(* IEC 61131-3 sources: plcassist-cli/packages/volt-lsp-iec/test-corpus/pro2193/Device/Plc Logic/Application/09 Misc/Library Manager/L_TS2P_TechModulesSynchronizingCamming (part 2) *)

(* ---- L_TS2P_SYNCANDCORRECTIONSTATE.fb ---- *)
FUNCTION_BLOCK L_TS2P_SYNCANDCORRECTIONSTATE EXTENDS L_TB2P_TechModuleBase
VAR_INPUT
	XUSEORIGINAL : BOOL;
	XENABLE : BOOL;
	XENABLEOPERATION : BOOL;
	XRESETERROR : BOOL;
	XQSPAPPLICATION : BOOL;
	XABORT : BOOL;
	XJOGPOS : BOOL;
	XJOGNEG : BOOL;
	XHOMEEXECUTE : BOOL;
	LROVERRIDE : LREAL := 1;
	SCCTRLBASICMOTION : L_TB2P_scCtrlBasicMotion;
	SCPAR : L_TS2P_scPar_SyncAndCorrectionState;
	SCACCESSPOINTS : L_TS2P_scAP_SyncAndCorrectionState;
	MASTERVALUES : L_MC1P_IAXIS_REF_MASTERVALUES;
	XSYNCIN : BOOL;
	XSYNCPOSRESTORE : BOOL;
	LRSETBASEVEL : LREAL;
	LRSETOFFSETPOS : LREAL;
	XTRIMPOS : BOOL;
	XTRIMNEG : BOOL;
	XTRIMRESET : BOOL;
	SCTPRECDATA_MARKSENSOR : L_MC1P_TpReceiveData;
	SCTPRECDATA_TOOLSENSOR : L_MC1P_TpReceiveData;
	XTEACHMARKWINDOW : BOOL;
	XTEACHMARKWINDOWTOOL : BOOL;
	XGEARFACTORCORR : BOOL;
	XGEARFACTORCORRHOLD : BOOL;
END_VAR
VAR_OUTPUT
	XREADYFOROPERATION : BOOL;
	XOPERATIONENABLED : BOOL;
	XREADYFORMOTION : BOOL;
	XERROR : BOOL;
	XWARNING : BOOL;
	EERRORID : L_IE1P_Error;
	XSTOACTIVE : BOOL;
	XQSPACTIVE : BOOL;
	XABORTBUSY : BOOL;
	XABORTDONE : BOOL;
	XJOGGINGBUSY : BOOL;
	XHOMINGBUSY : BOOL;
	XHOMINGDONE : BOOL;
	XISHOMED : BOOL;
	ETMSTATE : L_TB2P_States := L_TB2P_States.DISABLED;
	SCSTATUSBASICMOTION : L_TB2P_scStatusBasicMotion;
	LRACTVEL : LREAL;
	LRSETVELOUT : LREAL;
	LRACTPOS : LREAL;
	LRSETPOSOUT : LREAL;
	LRACTFOLLOWINGERROR : LREAL;
	SCSIGNALFLOW : L_TS2P_scSF_SyncAndCorrectionState;
	XSYNCHRONISED : BOOL;
	XACCDECSYNC : BOOL;
	XOFFSETTRIMACTIVE : BOOL;
	XBASEVELOCITYACTIVE : BOOL;
	LROFFSETTOTAL : LREAL;
	LRSETMARKCORROUT : LREAL;
	XMARKWINDOWTEACHED : BOOL;
	LRGEARFACTORCORR : LREAL;
	LRSETTOOLCORROUT : LREAL;
	XMARKWINDOWTEACHEDTOOL : BOOL;
END_VAR
VAR_IN_OUT
	AXIS : AXIS_REF;
END_VAR
VAR
	XINTERNALCONTROL : BOOL;
	XINTERNALCONTROLACTIVE : BOOL;
	XINTERNALCONTROLACTIVE_OLD : BOOL;
	ITFCONNECTORSYNCANDCORRECTION : L_TS2P_IConnectorSyncAndCorrection;
	TM_INT : L_TS2P_TM_SyncAndCorrectionState;
	SCPAR_INT : L_TS2P_scPar_SyncAndCorrectionState;
	XSYNCIN_INT : BOOL;
	XSYNCPOSRESTORE_INT : BOOL;
	LRSETBASEVEL_INT : LREAL;
	LRSETOFFSETPOS_INT : LREAL;
	XTRIMPOS_INT : BOOL;
	XTRIMNEG_INT : BOOL;
	XTRIMRESET_INT : BOOL;
	XTEACHMARKWINDOW_INT : BOOL;
	XTEACHMARKWINDOWTOOL_INT : BOOL;
	XGEARFACTORCORR_INT : BOOL;
	XGEARFACTORCORRHOLD_INT : BOOL;
	XUSEORIGINAL_OLD : BOOL;
	ITFBASICMOTIONBASE : L_TB2P.L_TB2P_IBasicMotionBase;
	ITFITECHMODULEINTERNAL : L_TB2P_ITechModuleInternal;
	ITFSYNCANDCORRECTIONEXTENSION : L_TS2P_ISyncAndCorrectionState;
	ITFSYNCPOSEXTENSION : L_TS2P_ISyncPosBase;
	LRJERKDEC : LREAL;
	LRJOGGINGJERKDEC : LREAL;
	REMAININGTIMEOFPROFILE : LREAL;
	REMAININGTIMEOFPROFILEAVAILABLE : BOOL;
END_VAR
END_FUNCTION_BLOCK

METHOD GET_PAP : POINTER TO L_TB2P_scAP_TM_MotionControl
END_METHOD

METHOD GET_PPAR : POINTER TO L_TB2P.L_TB2P_scPar_TM_MotionControl
END_METHOD

METHOD GET_PSF : POINTER TO L_TB2P_scSF_TM_MotionControl
END_METHOD

METHOD CALL_ABC
VAR_INPUT
	ITFTECHMODULE : L_TB2P.L_TB2P_IBasicMotionBase;
	XQSPAPPLICATION : BOOL;
	XHALT : BOOL;
	XABORT : BOOL;
	XHOMEEXECUTE : BOOL;
	XJOGPOS : BOOL;
	XJOGNEG : BOOL;
	XFINISHPOSITIONING : BOOL;
	XMOVEVELEXECUTE : BOOL;
	XMOVEABSEXECUTE : BOOL;
	XMOVERELEXECUTE : BOOL;
	XENABLEOPERATION : BOOL;
	XRESETERROR : BOOL;
	XENABLEPOSITIVE : BOOL;
	XENABLENEGATIVE : BOOL;
	XDISABLESWLIMIT : BOOL;
	LROVERRIDE : LREAL;
	LROVERRIDEACC : LREAL;
	LROVERRIDEJERK : LREAL;
	XRESETHOMEPOSITION : BOOL;
	XCONTINUOUSUPDATE : BOOL;
	LRPOS_DIST : LREAL;
	LRVEL : LREAL;
	LRACC : LREAL;
	LRDEC : LREAL;
	LRJERK : LREAL;
	EDIRECTION : L_TB2P.MC_DIRECTION;
	SCHOMEEXTTP : L_TB2P.MC_TRIGGER_REF;
	XHOMEABSSWITCH : BOOL;
	XSPECIALABORTBEHAVIOR : BOOL;
	LRABORTDEC : LREAL;
	LRABORTJERK : LREAL;
END_VAR
VAR_OUTPUT
	XERROR : BOOL;
	EERRORID : L_TB2P.L_IE1P_Error;
	XFUNBUSY : BOOL;
	XFUNDONE : BOOL;
	XFUNCOMMANDABORTED : BOOL;
	EFUNSTATEACT : L_TB2P.L_MC1P_ABC_State;
	ECONTROLMODE : L_TB2P.L_MC1P_ControlMode;
	XISHOMED : BOOL;
	XHWLIMITSWITCHNEG : BOOL;
	XHWLIMITSWITCHPOS : BOOL;
	XSWLIMITENABLED : BOOL;
	XSWLIMITSWITCHNEG : BOOL;
	XSWLIMITSWITCHPOS : BOOL;
	EAXISTYPE : L_TB2P.L_MC1P_DriveType;
	EAXISSTATE : L_TB2P.L_MC1P_AXIS_STATE;
	XSTOACTIVE : BOOL;
	XREADYFOROPERATION : BOOL;
	XOPERATIONENABLED : BOOL;
	XREADYFORMOTION : BOOL;
	XAXISWARNING : BOOL;
	XAXISERROR : BOOL;
	EAXISERRORID : L_TB2P.L_IE1P_Error;
	XDRIVEWARNING : BOOL;
	XDRIVEERROR : BOOL;
	DWDRIVEERRORID : DWORD;
	LRACTPOS : LREAL;
	LRACTVEL : LREAL;
	LRSETPOSOUT : LREAL;
	LRSETVELOUT : LREAL;
	LRACTFOLLOWINGERROR : LREAL;
	XINPOSITION : BOOL;
	XSTANDSTILLSETVELOCITY : BOOL;
	XSTANDSTILLACTVELOCITY : BOOL;
	XCONSTANTVELOCITY : BOOL;
	XACCELERATING : BOOL;
	XDECELERATING : BOOL;
	XDIRECTIONPOSITIVE : BOOL;
	XDIRECTIONNEGATIVE : BOOL;
	XAXISAVAILABLE : BOOL;
END_VAR
VAR_IN_OUT
	AXIS : AXIS_REF;
END_VAR
END_METHOD

METHOD ADDOFFSET
VAR_INPUT
	ITFTECHMODULE : L_TS2P_ISyncPosBase;
	LRSETPOS : LREAL;
	LRSETVEL : LREAL;
	LRSETOFFSET : LREAL;
	LRSETOFFSETVEL : LREAL;
	ETRAVERSINGRANGE : L_MC1P.L_MC1P_TraversingRange;
	LRCYCLELENGTH : LREAL;
END_VAR
VAR_OUTPUT
	XERROR : BOOL;
	EERRORID : L_IE1P.L_IE1P_Error;
	LRSETPOSOUT : LREAL;
	LRSETVELOUT : LREAL;
END_VAR
END_METHOD

METHOD CLUTCH
VAR_INPUT
	ITFTECHMODULE : L_TS2P_ISyncPosBase;
	XENABLE : BOOL;
	XSYNCIN : BOOL;
	LRSETBASEVELOCITY : LREAL;
	ESYNCMODE : L_TB2P_SyncMode;
	EALLOWEDDIRECTION : L_TB2P_AllowedDirection;
	LRSYNCVEL : LREAL;
	LRSYNCACC : LREAL;
	LRSYNCDEC : LREAL;
	LRSYNCJERK : LREAL;
	LRSYNCINDIST : LREAL;
	LRSYNCOUTDIST : LREAL;
	LRSYNCOUTPOS : LREAL;
	XLOADCLUTCHOFFSET : BOOL;
	LRLOADCLUTCHOFFSET : LREAL;
	LRCYCLICMASTERPOS : LREAL;
	LRCYCLICMASTERVEL : LREAL;
	ETRAVERSINGRANGEMASTER : L_MC1P_TraversingRange;
	LRCYCLELENGTHMASTER : LREAL;
	LRCYCLICAXISPOS : LREAL;
	LRCYCLICAXISVEL : LREAL;
	LRCYCLICAXISACC : LREAL;
	ETRAVERSINGRANGEAXIS : L_MC1P_TraversingRange;
	LRCYCLELENGTHAXIS : LREAL;
END_VAR
VAR_OUTPUT
	XERROR : BOOL;
	EERRORID : L_IE1P.L_IE1P_Error;
	XBUSY : BOOL;
	XDONE : BOOL;
	XSYNCHRONISED : BOOL;
	XACCDECSYNC : BOOL;
	XINBASEVELOCITY : BOOL;
	LRSETPOSOUT : LREAL;
	LRSETVELOUT : LREAL;
	LRSETACCOUT : LREAL;
	LRCLUTCHOFFSETOUT : LREAL;
END_VAR
END_METHOD

METHOD GEARBOX
VAR_INPUT
	ITFTECHMODULE : L_TS2P_ISyncPosBase;
	XENABLE : BOOL;
	LRSETPOSX : LREAL;
	LRSETVELX : LREAL;
	DWNUMERATOR : DWORD;
	DWDENOMINATOR : DWORD;
	LRCYCLELENGTHX : LREAL;
	LRCYCLELENGTHY : LREAL;
	ETRAVERSINGRANGEX : L_MC1P.L_MC1P_TraversingRange;
	ETRAVERSINGRANGEY : L_MC1P.L_MC1P_TraversingRange;
	XLOADGEARBOXPOS : BOOL;
	LRLOADGEARBOXPOS : LREAL;
END_VAR
VAR_OUTPUT
	XERROR : BOOL;
	EERRORID : L_IE1P.L_IE1P_Error;
	LRSETPOSOUT : LREAL;
	LRSETVELOUT : LREAL;
END_VAR
END_METHOD

METHOD OFFSETANDTRIM
VAR_INPUT
	ITFTECHMODULE : L_TS2P_ISyncPosBase;
	XENABLE : BOOL;
	LRSETOFFSET : LREAL;
	XTRIMPOS : BOOL;
	XTRIMNEG : BOOL;
	LRSETTRIMDISTANCE : LREAL;
	ETRIMMODE : L_TS2P_TrimMode;
	XLOADOFFSET : BOOL;
	XRESETTRIMOFFSET : BOOL;
	LRSETVEL : LREAL;
	LRSETACC : LREAL;
	LRSETDEC : LREAL;
	LRSETJERK : LREAL;
	WACTDIRECTION : WORD;
	EALLOWEDDIRECTION : L_TB2P.L_TB2P_AllowedDirection;
	LRCYCMASTERPOS : LREAL;
	LRCYCMASTERVEL : LREAL;
	LRCYCMASTERACC : LREAL;
END_VAR
VAR_OUTPUT
	XERROR : BOOL;
	EERRORID : L_IE1P.L_IE1P_Error;
	XBUSY : BOOL;
	XDONE : BOOL;
	LRSETOFFSETOUTTOTAL : LREAL;
	LRSETOFFSETOUTTOTALVEL : LREAL;
	LRSETOFFSETOUT : LREAL;
	LRSETOFFSETOUTTRIM : LREAL;
END_VAR
END_METHOD

METHOD FB_INIT : BOOL
VAR_INPUT
	BINITRETAINS : BOOL;
	BINCOPYCODE : BOOL;
END_VAR
END_METHOD

METHOD CALL_INTERNALCTRL
END_METHOD

(* ---- L_TS2P_SYNCANDCORRECTIONSTATE_V2.fb ---- *)
FUNCTION_BLOCK L_TS2P_SYNCANDCORRECTIONSTATE_V2 EXTENDS L_TB2P_TechModuleBase
VAR_INPUT
	XENABLE : BOOL;
	XENABLEOPERATION : BOOL;
	XRESETERROR : BOOL;
	XQSPAPPLICATION : BOOL;
	XABORT : BOOL;
	XJOGPOS : BOOL;
	XJOGNEG : BOOL;
	XHOMEEXECUTE : BOOL;
	LROVERRIDE : LREAL := 1;
	SCCTRLBASICMOTION : L_TB2P_scCtrlBasicMotion;
	SCPAR : L_TS2P_scPar_SyncAndCorrectionState;
	SCACCESSPOINTS : L_TS2P_scAP_SyncAndCorrectionState;
	MASTERVALUES : L_MC1P_IAXIS_REF_MASTERVALUES;
	XSYNCIN : BOOL;
	XSYNCPOSRESTORE : BOOL;
	LRSETBASEVEL : LREAL;
	LRSETOFFSETPOS : LREAL;
	XTRIMPOS : BOOL;
	XTRIMNEG : BOOL;
	XTRIMRESET : BOOL;
	SCTPRECDATA_MARKSENSOR : L_MC1P_TpReceiveData;
	SCTPRECDATA_TOOLSENSOR : L_MC1P_TpReceiveData;
	XTEACHMARKWINDOW : BOOL;
	XTEACHMARKWINDOWTOOL : BOOL;
	XGEARFACTORCORR : BOOL;
	XGEARFACTORCORRHOLD : BOOL;
END_VAR
VAR_OUTPUT
	XREADYFOROPERATION : BOOL;
	XOPERATIONENABLED : BOOL;
	XREADYFORMOTION : BOOL;
	XERROR : BOOL;
	XWARNING : BOOL;
	EERRORID : L_IE1P_Error;
	XSTOACTIVE : BOOL;
	XQSPACTIVE : BOOL;
	XABORTBUSY : BOOL;
	XABORTDONE : BOOL;
	XJOGGINGBUSY : BOOL;
	XHOMINGBUSY : BOOL;
	XHOMINGDONE : BOOL;
	XISHOMED : BOOL;
	ETMSTATE : L_TB2P_States := L_TB2P_States.DISABLED;
	SCSTATUSBASICMOTION : L_TB2P_scStatusBasicMotion;
	LRACTVEL : LREAL;
	LRSETVELOUT : LREAL;
	LRACTPOS : LREAL;
	LRSETPOSOUT : LREAL;
	LRACTFOLLOWINGERROR : LREAL;
	SCSIGNALFLOW : L_TS2P_scSF_SyncAndCorrectionState;
	XSYNCHRONISED : BOOL;
	XACCDECSYNC : BOOL;
	XOFFSETTRIMACTIVE : BOOL;
	XBASEVELOCITYACTIVE : BOOL;
	LROFFSETTOTAL : LREAL;
	LRSETMARKCORROUT : LREAL;
	XMARKWINDOWTEACHED : BOOL;
	LRGEARFACTORCORR : LREAL;
	LRSETTOOLCORROUT : LREAL;
	XMARKWINDOWTEACHEDTOOL : BOOL;
END_VAR
VAR_IN_OUT
	AXIS : AXIS_REF;
END_VAR
VAR
	TM_INT : L_TS2P_TM_SyncAndCorrectionState_V2 := STRUCT(ModuleHandler := ModuleHandler);
	PPAR : POINTER TO L_TS2P_scPar_SyncAndCorrectionState;
	PPAR_INT : POINTER TO L_TS2P_scPar_SyncAndCorrectionState;
	LRJERKDEC : LREAL;
	LRJOGGINGJERKDEC : LREAL;
END_VAR
END_FUNCTION_BLOCK

(* ---- L_TS2P_SYNCDRIVEPOS.fb ---- *)
FUNCTION_BLOCK L_TS2P_SYNCDRIVEPOS
VAR_INPUT
	MASTERAXIS : POINTER TO L_MC1P_IAXIS_REF_MASTERVALUES;
	XENABLE : BOOL;
	DWNUMERATOR : DWORD := 1;
	DWDENOMINATOR : DWORD := 1;
	XSYNCIN : BOOL;
	XSYNCOUTINSTANT : BOOL;
	XSYNCINSTANT : BOOL;
	XCLUTCHRELATIVE : BOOL;
	XSYNCPOSRESTORE : BOOL;
	LRSLAVESYNCOUTPOS : LREAL;
	LRSLAVESYNCINDIST : LREAL := 90;
	LRSLAVESYNCOUTDIST : LREAL := 90;
	LRSYNCOUTINSTANTDEC : LREAL := 10000;
	EALLOWEDDIRECTION : L_TB2P_AllowedDirection := L_TB2P_AllowedDirection.both;
	ESYNCMODE : L_TB2P_SyncMode := L_TB2P_SyncMode.ProfGenAbsolute;
	LRSYNCVEL : LREAL := 100;
	LRSYNCACC : LREAL := 1000.0;
	LRSYNCDEC : LREAL := 1000.0;
	LRSYNCJERK : LREAL := 10000000000.0;
	LRSETBASEVELOCITY : LREAL := 0;
	XLOADCLUTCHOFFSET : BOOL := FALSE;
	LRLOADCLUTCHOFFSET : LREAL := 0;
	XTRIMVELOCITYX : BOOL;
	XTRIMVELOCITYY : BOOL;
	LRSETTRIMDISTANCEX : LREAL := 1;
	LRSETTRIMDISTANCEY : LREAL := 1;
	XTRIMPOSX : BOOL;
	XTRIMNEGX : BOOL;
	XTRIMPOSY : BOOL;
	XTRIMNEGY : BOOL;
	XRESETTRIMX : BOOL;
	XRESETTRIMY : BOOL;
	LRSETOFFSETX : LREAL := 0;
	LRSETOFFSETTRIMVELX : LREAL := 10.0;
	LRSETOFFSETTRIMACCX : LREAL := 100.0;
	LRSETOFFSETTRIMDECX : LREAL := 100.0;
	LRSETOFFSETTRIMJERKX : LREAL := 10000.0;
	XLOADOFFSETX : BOOL;
	LRSETOFFSETY : LREAL := 0;
	LRSETOFFSETTRIMVELY : LREAL := 10.0;
	LRSETOFFSETTRIMACCY : LREAL := 100.0;
	LRSETOFFSETTRIMDECY : LREAL := 100.0;
	LRSETOFFSETTRIMJERKY : LREAL := 10000.0;
	XLOADOFFSETY : BOOL;
	XLOADSTARTSLAVEPOS : BOOL := FALSE;
	LRSTARTSLAVEPOS : LREAL;
	XLOADGEARBOXPOS : BOOL;
	LRLOADGEARBOXPOS : LREAL;
	XOPERATIONENABLED : BOOL;
END_VAR
VAR_OUTPUT
	XERROR : BOOL;
	XWARNING : BOOL;
	EERRORID : L_IE1P_Error;
	XBUSY : BOOL;
	LRSETSLAVEPOSOUT : LREAL;
	LRSETSLAVEVELOUT : LREAL;
	LRSETSLAVEACCOUT : LREAL;
	LRSETGEARBOXPOSOUT : LREAL;
	XSYNCOUTDONE : BOOL;
	XSYNCHRONISED : BOOL;
	XACCDECSYNC : BOOL;
	XOFFSETTRIMBUSY : BOOL;
	LROFFSETOUTTOTALVELX : LREAL;
	LROFFSETOUTTOTALVELY : LREAL;
	LROFFSETOUTTRIMX : LREAL;
	LROFFSETOUTTRIMY : LREAL;
	LROFFSETOUTX : LREAL;
	LROFFSETOUTY : LREAL;
	LROFFSETOUTTOTALX : LREAL;
	LROFFSETOUTTOTALY : LREAL;
	LRSETCLUTCHPOS : LREAL;
	LRSETCLUTCHVEL : LREAL;
	LRSETCLUTCHACC : LREAL;
	XBASEVELSYNCHRONISED : BOOL;
	XACCDECBASEVEL : BOOL;
	LROFFSETSYNCPOS : LREAL;
END_VAR
VAR_IN_OUT
	SLAVEAXIS : AXIS_REF;
END_VAR
VAR
	FB_GEARBOXPOSITION : L_MB1P_GearboxPositionInput;
	FB_CLUTCHEXTENDEDBASE : L_TB2P_ClutchExtendedBase;
	FB_AXISCONVERTER : L_MC2P.L_MC2P_AxisConverterBase;
	FB_OFFSETANDTRIMX : L_TS2P_OffsetAndTrim;
	FB_ADDOFFSETCYCLICX : L_MC1P_AddOffsetCyclic;
	FB_OFFSETANDTRIMY : L_TS2P_OffsetAndTrim;
	FB_ADDOFFSETCYCLICY : L_MC1P_AddOffsetCyclic;
	FB_SYNCPOSRESTOREOFFSET : L_TS2P_OffsetAndTrim;
	FB_DIRECTION : L_MC1P_GetDirection;
	LRSETOFFSETMASTER_INT : LREAL;
	LRTRIMDIST_INT : LREAL;
	XTRIMPOS_OLD : BOOL;
	XTRIMNEG_OLD : BOOL;
	XTRIMVEL : BOOL;
	LRTRIMOFFSETDIST : LREAL;
	LRLOADOFFSETMASTER_INT : LREAL := 0;
	LRLOADGEARBOXPOS_INT : LREAL;
	LRSETGEARBOXPOSOUT_INT : LREAL;
	XSETDISABLECLUTCH_INT : BOOL;
	LRLOADTRIMOFFSET_INT : LREAL := 0;
	LRSYNCOUTINSTANTDEC_INT : LREAL := 100000;
	LRSETINTEGRATETRIMVELPOSOUT_INT : LREAL;
	XSYNCPOS_OLD : BOOL;
	XRESETTRIM_OLD : BOOL;
	LRLOADOFFSET_INT : LREAL := 0;
	XSYNCINSTANT_OLD : BOOL;
	XENABLEGEARBOX : BOOL;
	LRSYNCOFFSET : LREAL;
	LRSCALING_INT : LREAL := 1;
	LRGEARBOXSTARTPOSOUT_INT : LREAL;
	DWDENOMINATOR_INT : DWORD := 1;
	XENABLE_OLD : BOOL;
	WAXESMODE : WORD;
	WAXESMODEOLD : WORD;
	LRADDOFFSETPOSOUTY_OLD : LREAL;
	LRADDOFFSETVELOUTY : LREAL;
	LRSETGEARBOXPOSOUTOLD_INT : LREAL;
	LRSETGEARBOXPOSOUTVEL_INT : LREAL;
	LRGETGEARBOXVELIN : LREAL;
	LRGETGEARBOXPOSOUT : LREAL;
	LRGETGEARBOXPOSIN : LREAL;
	LRTASKCYCLE : LREAL;
	XINIT : BOOL := TRUE;
	XCLUTCHDONE_OLD : BOOL;
	XENABLEOLD : BOOL;
	LRSETOFFSETOUTTOTALVELOLD : LREAL;
	SET_AP_LRMASTERVELSTANDSTILLDEADBAND : LREAL;
END_VAR
END_FUNCTION_BLOCK

METHOD CALL_AXESMODE
END_METHOD

METHOD CALL_CALCGEARBOXOUTVELACC
VAR_IN_OUT
	SLAVEAXIS : AXIS_REF;
END_VAR
END_METHOD

METHOD CALL_ERRORHANDLER
END_METHOD

METHOD CALL_FBMETHODS
END_METHOD

METHOD CALL_FBMETHODS_FMDISABLE
END_METHOD

METHOD CALL_FB_ADDOFFSETCYCLICX
END_METHOD

METHOD CALL_FB_ADDOFFSETCYCLICX_INPUT
END_METHOD

METHOD CALL_FB_ADDOFFSETCYCLICY
END_METHOD

METHOD CALL_FB_ADDOFFSETCYCLICY_INPUT
END_METHOD

METHOD CALL_FB_AXISCONVERTER
END_METHOD

METHOD CALL_FB_AXISCONVERTER_INPUT
END_METHOD

METHOD CALL_FB_CLUTCHEXTENDEDBASE
END_METHOD

METHOD CALL_FB_CLUTCHEXTENDEDBASE_INPUT
END_METHOD

METHOD CALL_FB_CLUTCHEXTENDEDBASE_INPUTMASTER
END_METHOD

METHOD CALL_FB_CLUTCHEXTENDEDBASE_INPUTSLAVE
VAR_IN_OUT
	SLAVEAXIS : AXIS_REF;
END_VAR
END_METHOD

METHOD CALL_FB_GEARBOXPOSITION
END_METHOD

METHOD CALL_FB_GEARBOXPOSITION_INPUT
END_METHOD

METHOD CALL_FB_GEARBOXPOSITION_LOADGEARBOXPOS
END_METHOD

METHOD CALL_FB_SYNCPOSRESTOREOFFSET
END_METHOD

METHOD CALL_FB_SYNCPOSRESTOREOFFSET_INPUT
VAR_IN_OUT
	SLAVEAXIS : AXIS_REF;
END_VAR
END_METHOD

METHOD CALL_LOADSLAVESTARTPOS
END_METHOD

METHOD CALL_OFFSETANDTRIMX
END_METHOD

METHOD CALL_OFFSETANDTRIMX_INPUT
END_METHOD

METHOD CALL_OFFSETANDTRIMY
END_METHOD

METHOD CALL_OFFSETANDTRIMY_INPUT
END_METHOD

METHOD CALL_OUTPUT
END_METHOD

METHOD CALL_OUTPUT_CLUTCHSTATE
END_METHOD

METHOD CALL_OUTPUT_OFFSET
END_METHOD

METHOD CALL_RESETCOMMANDS
END_METHOD

METHOD CALL_INIT
VAR_IN_OUT
	SLAVEAXIS : AXIS_REF;
END_VAR
END_METHOD

METHOD GET_DIRECTION
END_METHOD

METHOD GET_GETGEARBOXPOSIN : LREAL
END_METHOD

METHOD GET_GETGEARBOXPOSOUT : LREAL
END_METHOD

METHOD GET_GETGEARBOXVELIN : LREAL
END_METHOD

METHOD GET_GETGEARBOXVELOUT : LREAL
END_METHOD

METHOD GET_LRCLUTCHPOSIN : LREAL
END_METHOD

METHOD GET_LROFFSETADDOFFSETCYCLIC : LREAL
END_METHOD

METHOD SETDISABLECLUTCH : BOOL
VAR_INPUT
	XSETDISABLECLUTCH : BOOL;
END_VAR
END_METHOD

(* ---- L_TS2P_SYNCDRIVEVEL.fb ---- *)
FUNCTION_BLOCK L_TS2P_SYNCDRIVEVEL
VAR_INPUT
	MASTERAXIS : POINTER TO L_MC1P_IAXIS_REF_MASTERVALUES;
	XENABLE : BOOL;
	LRCOUPLINGX : LREAL := 1.0;
	LRCOUPLINGY : LREAL := 1.0;
	XINVERTGEARFACTOR : BOOL;
	XDISABLETOLERANCEINVERTGEARFACTOR : BOOL;
	LRTOLERANCEINVERTGEARFACTOR : LREAL := 0;
	XSYNCIN : BOOL;
	XSYNCOUTINSTANT : BOOL;
	LRSYNCACC : LREAL := 10.0;
	LRSYNCDEC : LREAL := 10.0;
	LRSYNCOUTINSTANTDEC : LREAL := 100.0;
	LRSYNCJERK : LREAL := 1.0;
	XAVOIDVELGAPS : BOOL;
	LRSETOFFSETVEL : LREAL;
	DWMODE : DWORD := 1;
	XTRIMVELOCITYX : BOOL;
	XTRIMVELOCITYY : BOOL;
	LRSETTRIMDISTANCEX : LREAL := 1;
	LRSETTRIMDISTANCEY : LREAL := 1;
	XTRIMPOSX : BOOL;
	XTRIMNEGX : BOOL;
	XTRIMPOSY : BOOL;
	XTRIMNEGY : BOOL;
	XRESETTRIMX : BOOL;
	XRESETTRIMY : BOOL;
	XSYNCVELRESET : BOOL;
	LRSETOFFSETX : LREAL := 0;
	LRSETOFFSETTRIMVELX : LREAL := 10.0;
	LRSETOFFSETTRIMACCX : LREAL := 100.0;
	LRSETOFFSETTRIMDECX : LREAL := 100.0;
	LRSETOFFSETTRIMJERKX : LREAL := 10000.0;
	XLOADOFFSETX : BOOL;
	LRSETOFFSETY : LREAL := 0;
	LRSETOFFSETTRIMVELY : LREAL := 10.0;
	LRSETOFFSETTRIMACCY : LREAL := 100.0;
	LRSETOFFSETTRIMDECY : LREAL := 100.0;
	LRSETOFFSETTRIMJERKY : LREAL := 10000.0;
	XLOADOFFSETY : BOOL;
	EALLOWEDDIRECTION : L_TB2P_AllowedDirection;
	XLOADOFFSET : BOOL;
	XLOADGROUNDVEL : BOOL;
	LRSETGROUNDVEL : LREAL;
	LRGROUNDVELACC : LREAL := 10.0;
	LRGROUNDVELDEC : LREAL := 10.0;
	LRGROUNDVELJERK : LREAL := 1.0;
END_VAR
VAR_OUTPUT
	XERROR : BOOL;
	XWARNING : BOOL;
	EERRORID : L_IE1P_Error;
	XBUSY : BOOL;
	LRSETSLAVEVELOUT : LREAL;
	LRSETSLAVEACCOUT : LREAL;
	XSYNCOUTDONE : BOOL;
	XSYNCHRONISED : BOOL;
	XACCDECSYNC : BOOL;
	XOFFSETTRIMBUSY : BOOL;
	LRPOSOFFSETOUTTRIMX : LREAL;
	LRPOSOFFSETOUTTRIMY : LREAL;
	LRPOSOFFSETOUTX : LREAL;
	LRPOSOFFSETOUTY : LREAL;
	LRPOSOFFSETOUTVELX : LREAL;
	LRVELOFFSET : LREAL;
	LROFFSETOUTTOTALX : LREAL;
	LROFFSETOUTTOTALY : LREAL;
	LROFFSETOUTTOTALVELX : LREAL;
	LROFFSETOUTTOTALVELY : LREAL;
	XBASEVELSYNCHRONISED : BOOL;
	XACCDECBASEVEL : BOOL;
	XBASEVELSYNCOUTDONE : BOOL;
	XINVERTGEARFACTORACTIVE : BOOL;
END_VAR
VAR_IN_OUT
	SLAVEAXIS : AXIS_REF;
END_VAR
VAR
	XENABLE_OLD : BOOL;
	ESTATE : L_TF1P_States := L_TF1P_States.INIT;
	ESTATE_OLD : L_TF1P_States := L_TF1P_States.INIT;
	XSTATEENTRY : BOOL;
	FB_CONVAXISV : L_MC2P_ConvAxisV;
	FB_INVERTGEARFACTOR : L_TS2P_InvertGearfactor;
	XACCDECSYNC_OLD : BOOL;
	XSYNCVEL_OLD : BOOL;
	XOPEN_OLD : BOOL;
	LRSETVELTRIM : LREAL;
	XSETDISABLECLUTCH_INT : BOOL;
	SETPOSITIONFORSYNCOLD : LREAL := 0;
	XINITFB_CLUTCHV : BOOL;
	FB_CLUTCHV : L_MC2P_ClutchVelocity;
	XINVERTGEARFACTORACTIVE_OLD : BOOL;
	LRSETGROUNDVEL_INT : LREAL;
	FB_OFFSETANDTRIMX : L_TS2P_OffsetAndTrim;
	FB_VELOCITYOFFSET : L_MC1P_RampGenerator;
	FB_OFFSETANDTRIMY : L_TS2P_OffsetAndTrim;
	FB_RAMPGENGROUNDVEL : L_MC1P_RampGenerator;
	FB_DIRECTION : L_MC1P_GetDirection;
END_VAR
END_FUNCTION_BLOCK

METHOD CALL_ERRORHANDLER
END_METHOD

METHOD CALL_FBMETHODS
END_METHOD

METHOD CALL_FBMETHODS_FMDISABLE
END_METHOD

METHOD CALL_FB_CLUTCHV
END_METHOD

METHOD CALL_FB_CLUTCHV_INPUT
END_METHOD

METHOD CALL_FB_CLUTCHV_PAR
END_METHOD

METHOD CALL_FB_CONVAXISV
END_METHOD

METHOD CALL_FB_CONVAXISV_INPUT
END_METHOD

METHOD CALL_FB_INVERTGEARFACTOR
END_METHOD

METHOD CALL_FB_INVERTGEARFACTOR_INPUT
END_METHOD

METHOD CALL_FB_RAMPGENGROUNDVEL
END_METHOD

METHOD CALL_FB_RAMPGENGROUNDVEL_INPUT
END_METHOD

METHOD CALL_FB_VELOCITYOFFSET
END_METHOD

METHOD CALL_FB_VELOCITYOFFSET_INPUT
END_METHOD

METHOD CALL_OFFSETANDTRIMX
END_METHOD

METHOD CALL_OFFSETANDTRIMX_INPUT
END_METHOD

METHOD CALL_OFFSETANDTRIMY
END_METHOD

METHOD CALL_OFFSETANDTRIMY_INPUT
END_METHOD

METHOD CALL_OUTPUT
END_METHOD

METHOD CALL_OUTPUT_SETSLAVEOUT
END_METHOD

METHOD CALL_RESETCOMMANDS
END_METHOD

METHOD CALL_RESETFM
END_METHOD

METHOD CALL_RESETOUTPUT
END_METHOD

METHOD CALL_STATEMASHINE
END_METHOD

METHOD GET_DIRECTION
END_METHOD

METHOD GET_CLUTCHVELOUT : LREAL
END_METHOD

METHOD GET_GETGEARBOXVELIN : LREAL
END_METHOD

METHOD GET_GETGEARBOXVELOUT : LREAL
END_METHOD

METHOD SETDISABLECLUTCH : BOOL
VAR_INPUT
	XSETDISABLECLUTCH : BOOL;
END_VAR
END_METHOD

METHOD CALL_S000_CYCLIC
END_METHOD

METHOD CALL_S001_INIT
END_METHOD

METHOD CALL_S010_READY
END_METHOD

METHOD CALL_S998_ERROR
END_METHOD

(* ---- L_TS2P_SYNCPOSBASE.fb ---- *)
FUNCTION_BLOCK L_TS2P_SYNCPOSBASE EXTENDS L_TB2P_TechModuleBase
VAR_INPUT
	XUSEORIGINAL : BOOL;
	XENABLE : BOOL;
	XENABLEOPERATION : BOOL;
	XRESETERROR : BOOL;
	XQSPAPPLICATION : BOOL;
	XABORT : BOOL;
	XJOGPOS : BOOL;
	XJOGNEG : BOOL;
	XHOMEEXECUTE : BOOL;
	LROVERRIDE : LREAL := 1;
	SCCTRLBASICMOTION : L_TB2P_scCtrlBasicMotion;
	SCPAR : L_TS2P_scPar_SyncPosBase;
	SCACCESSPOINTS : L_TS2P_scAP_SyncPosBase;
	MASTERVALUES : L_MC1P_IAXIS_REF_MASTERVALUES;
	XSYNCIN : BOOL;
	XSYNCPOSRESTORE : BOOL;
	LRSETBASEVEL : LREAL;
	LRSETOFFSETPOS : LREAL;
	XTRIMPOS : BOOL;
	XTRIMNEG : BOOL;
	XTRIMRESET : BOOL;
END_VAR
VAR_OUTPUT
	XREADYFOROPERATION : BOOL;
	XOPERATIONENABLED : BOOL;
	XREADYFORMOTION : BOOL;
	XERROR : BOOL;
	XWARNING : BOOL;
	EERRORID : L_IE1P_Error;
	XSTOACTIVE : BOOL;
	XQSPACTIVE : BOOL;
	XABORTBUSY : BOOL;
	XABORTDONE : BOOL;
	XJOGGINGBUSY : BOOL;
	XHOMINGBUSY : BOOL;
	XHOMINGDONE : BOOL;
	XISHOMED : BOOL;
	ETMSTATE : L_TB2P_States;
	SCSTATUSBASICMOTION : L_TB2P_scStatusBasicMotion;
	LRACTVEL : LREAL;
	LRSETVELOUT : LREAL;
	LRACTPOS : LREAL;
	LRSETPOSOUT : LREAL;
	LRACTFOLLOWINGERROR : LREAL;
	SCSIGNALFLOW : L_TS2P_scSF_SyncPosBase;
	XSYNCHRONISED : BOOL;
	XACCDECSYNC : BOOL;
	XOFFSETTRIMACTIVE : BOOL;
	XBASEVELOCITYACTIVE : BOOL;
	LROFFSETTOTAL : LREAL;
END_VAR
VAR_IN_OUT
	AXIS : AXIS_REF;
END_VAR
VAR
	XINTERNALCONTROL : BOOL;
	XINTERNALCONTROLACTIVE : BOOL;
	XINTERNALCONTROLACTIVE_OLD : BOOL;
	ITFCONNECTORSYNCPOS : L_TS2P_IConnectorSyncPos;
	TM_INT : L_TS2P_TM_SyncPosBase;
	SCPAR_INT : L_TS2P_scPar_SyncPosBase;
	XSYNCIN_INT : BOOL;
	XSYNCPOSRESTORE_INT : BOOL;
	LRSETBASEVEL_INT : LREAL;
	LRSETOFFSETPOS_INT : LREAL;
	LRSETOFFSETVEL_INT : LREAL;
	XTRIMPOS_INT : BOOL;
	XTRIMNEG_INT : BOOL;
	XTRIMRESET_INT : BOOL;
	SCSIGNALFLOW_INT : L_TS2P_scSF_SyncPosBase;
	XUSEORIGINAL_OLD : BOOL;
	ITFBASICMOTIONBASE : L_TB2P.L_TB2P_IBasicMotionBase;
	ITFITECHMODULEINTERNAL : L_TB2P_ITechModuleInternal;
	ITFSYNCPOSEXTENSION : L_TS2P_ISyncPosBase;
	LRJERKDEC : LREAL;
	LRJOGGINGJERKDEC : LREAL;
	REMAININGTIMEOFPROFILE : LREAL;
	REMAININGTIMEOFPROFILEAVAILABLE : BOOL;
END_VAR
END_FUNCTION_BLOCK

METHOD GET_PAP : POINTER TO L_TB2P_scAP_TM_MotionControl
END_METHOD

METHOD GET_PPAR : POINTER TO L_TB2P.L_TB2P_scPar_TM_MotionControl
END_METHOD

METHOD GET_PSF : POINTER TO L_TB2P_scSF_TM_MotionControl
END_METHOD

METHOD CALL_ABC
VAR_INPUT
	ITFTECHMODULE : L_TB2P.L_TB2P_IBasicMotionBase;
	XQSPAPPLICATION : BOOL;
	XHALT : BOOL;
	XABORT : BOOL;
	XHOMEEXECUTE : BOOL;
	XJOGPOS : BOOL;
	XJOGNEG : BOOL;
	XFINISHPOSITIONING : BOOL;
	XMOVEVELEXECUTE : BOOL;
	XMOVEABSEXECUTE : BOOL;
	XMOVERELEXECUTE : BOOL;
	XENABLEOPERATION : BOOL;
	XRESETERROR : BOOL;
	XENABLEPOSITIVE : BOOL;
	XENABLENEGATIVE : BOOL;
	XDISABLESWLIMIT : BOOL;
	LROVERRIDE : LREAL;
	LROVERRIDEACC : LREAL;
	LROVERRIDEJERK : LREAL;
	XRESETHOMEPOSITION : BOOL;
	XCONTINUOUSUPDATE : BOOL;
	LRPOS_DIST : LREAL;
	LRVEL : LREAL;
	LRACC : LREAL;
	LRDEC : LREAL;
	LRJERK : LREAL;
	EDIRECTION : L_TB2P.MC_DIRECTION;
	SCHOMEEXTTP : L_TB2P.MC_TRIGGER_REF;
	XHOMEABSSWITCH : BOOL;
	XSPECIALABORTBEHAVIOR : BOOL;
	LRABORTDEC : LREAL;
	LRABORTJERK : LREAL;
END_VAR
VAR_OUTPUT
	XERROR : BOOL;
	EERRORID : L_TB2P.L_IE1P_Error;
	XFUNBUSY : BOOL;
	XFUNDONE : BOOL;
	XFUNCOMMANDABORTED : BOOL;
	EFUNSTATEACT : L_TB2P.L_MC1P_ABC_State;
	ECONTROLMODE : L_TB2P.L_MC1P_ControlMode;
	XISHOMED : BOOL;
	XHWLIMITSWITCHNEG : BOOL;
	XHWLIMITSWITCHPOS : BOOL;
	XSWLIMITENABLED : BOOL;
	XSWLIMITSWITCHNEG : BOOL;
	XSWLIMITSWITCHPOS : BOOL;
	EAXISTYPE : L_TB2P.L_MC1P_DriveType;
	EAXISSTATE : L_TB2P.L_MC1P_AXIS_STATE;
	XSTOACTIVE : BOOL;
	XREADYFOROPERATION : BOOL;
	XOPERATIONENABLED : BOOL;
	XREADYFORMOTION : BOOL;
	XAXISWARNING : BOOL;
	XAXISERROR : BOOL;
	EAXISERRORID : L_TB2P.L_IE1P_Error;
	XDRIVEWARNING : BOOL;
	XDRIVEERROR : BOOL;
	DWDRIVEERRORID : DWORD;
	LRACTPOS : LREAL;
	LRACTVEL : LREAL;
	LRSETPOSOUT : LREAL;
	LRSETVELOUT : LREAL;
	LRACTFOLLOWINGERROR : LREAL;
	XINPOSITION : BOOL;
	XSTANDSTILLSETVELOCITY : BOOL;
	XSTANDSTILLACTVELOCITY : BOOL;
	XCONSTANTVELOCITY : BOOL;
	XACCELERATING : BOOL;
	XDECELERATING : BOOL;
	XDIRECTIONPOSITIVE : BOOL;
	XDIRECTIONNEGATIVE : BOOL;
	XAXISAVAILABLE : BOOL;
END_VAR
VAR_IN_OUT
	AXIS : AXIS_REF;
END_VAR
END_METHOD

METHOD ADDOFFSET
VAR_INPUT
	ITFTECHMODULE : L_TS2P_ISyncPosBase;
	LRSETPOS : LREAL;
	LRSETVEL : LREAL;
	LRSETOFFSET : LREAL;
	LRSETOFFSETVEL : LREAL;
	ETRAVERSINGRANGE : L_MC1P.L_MC1P_TraversingRange;
	LRCYCLELENGTH : LREAL;
END_VAR
VAR_OUTPUT
	XERROR : BOOL;
	EERRORID : L_IE1P.L_IE1P_Error;
	LRSETPOSOUT : LREAL;
	LRSETVELOUT : LREAL;
END_VAR
END_METHOD

METHOD CLUTCH
VAR_INPUT
	ITFTECHMODULE : L_TS2P_ISyncPosBase;
	XENABLE : BOOL;
	XSYNCIN : BOOL;
	LRSETBASEVELOCITY : LREAL;
	ESYNCMODE : L_TB2P_SyncMode;
	EALLOWEDDIRECTION : L_TB2P_AllowedDirection;
	LRSYNCVEL : LREAL;
	LRSYNCACC : LREAL;
	LRSYNCDEC : LREAL;
	LRSYNCJERK : LREAL;
	LRSYNCINDIST : LREAL;
	LRSYNCOUTDIST : LREAL;
	LRSYNCOUTPOS : LREAL;
	XLOADCLUTCHOFFSET : BOOL;
	LRLOADCLUTCHOFFSET : LREAL;
	LRCYCLICMASTERPOS : LREAL;
	LRCYCLICMASTERVEL : LREAL;
	ETRAVERSINGRANGEMASTER : L_MC1P_TraversingRange;
	LRCYCLELENGTHMASTER : LREAL;
	LRCYCLICAXISPOS : LREAL;
	LRCYCLICAXISVEL : LREAL;
	LRCYCLICAXISACC : LREAL;
	ETRAVERSINGRANGEAXIS : L_MC1P_TraversingRange;
	LRCYCLELENGTHAXIS : LREAL;
END_VAR
VAR_OUTPUT
	XERROR : BOOL;
	EERRORID : L_IE1P.L_IE1P_Error;
	XBUSY : BOOL;
	XDONE : BOOL;
	XSYNCHRONISED : BOOL;
	XACCDECSYNC : BOOL;
	XINBASEVELOCITY : BOOL;
	LRSETPOSOUT : LREAL;
	LRSETVELOUT : LREAL;
	LRSETACCOUT : LREAL;
	LRCLUTCHOFFSETOUT : LREAL;
END_VAR
END_METHOD

METHOD GEARBOX
VAR_INPUT
	ITFTECHMODULE : L_TS2P_ISyncPosBase;
	XENABLE : BOOL;
	LRSETPOSX : LREAL;
	LRSETVELX : LREAL;
	DWNUMERATOR : DWORD;
	DWDENOMINATOR : DWORD;
	LRCYCLELENGTHX : LREAL;
	LRCYCLELENGTHY : LREAL;
	ETRAVERSINGRANGEX : L_MC1P.L_MC1P_TraversingRange;
	ETRAVERSINGRANGEY : L_MC1P.L_MC1P_TraversingRange;
	XLOADGEARBOXPOS : BOOL;
	LRLOADGEARBOXPOS : LREAL;
END_VAR
VAR_OUTPUT
	XERROR : BOOL;
	EERRORID : L_IE1P.L_IE1P_Error;
	LRSETPOSOUT : LREAL;
	LRSETVELOUT : LREAL;
END_VAR
END_METHOD

METHOD OFFSETANDTRIM
VAR_INPUT
	ITFTECHMODULE : L_TS2P_ISyncPosBase;
	XENABLE : BOOL;
	LRSETOFFSET : LREAL;
	XTRIMPOS : BOOL;
	XTRIMNEG : BOOL;
	LRSETTRIMDISTANCE : LREAL;
	ETRIMMODE : L_TS2P_TrimMode;
	XLOADOFFSET : BOOL;
	XRESETTRIMOFFSET : BOOL;
	LRSETVEL : LREAL;
	LRSETACC : LREAL;
	LRSETDEC : LREAL;
	LRSETJERK : LREAL;
	WACTDIRECTION : WORD;
	EALLOWEDDIRECTION : L_TB2P.L_TB2P_AllowedDirection;
	LRCYCMASTERPOS : LREAL;
	LRCYCMASTERVEL : LREAL;
	LRCYCMASTERACC : LREAL;
END_VAR
VAR_OUTPUT
	XERROR : BOOL;
	EERRORID : L_IE1P.L_IE1P_Error;
	XBUSY : BOOL;
	XDONE : BOOL;
	LRSETOFFSETOUTTOTAL : LREAL;
	LRSETOFFSETOUTTOTALVEL : LREAL;
	LRSETOFFSETOUT : LREAL;
	LRSETOFFSETOUTTRIM : LREAL;
END_VAR
END_METHOD

METHOD FB_INIT : BOOL
VAR_INPUT
	BINITRETAINS : BOOL;
	BINCOPYCODE : BOOL;
END_VAR
END_METHOD

METHOD CALL_INTERNALCTRL
END_METHOD

(* ---- L_TS2P_SYNCPOSBASE_V2.fb ---- *)
FUNCTION_BLOCK L_TS2P_SYNCPOSBASE_V2 EXTENDS L_TB2P_TechModuleBase
VAR_INPUT
	XENABLE : BOOL;
	XENABLEOPERATION : BOOL;
	XRESETERROR : BOOL;
	XQSPAPPLICATION : BOOL;
	XABORT : BOOL;
	XJOGPOS : BOOL;
	XJOGNEG : BOOL;
	XHOMEEXECUTE : BOOL;
	LROVERRIDE : LREAL := 1;
	SCCTRLBASICMOTION : L_TB2P_scCtrlBasicMotion;
	SCPAR : L_TS2P_scPar_SyncPosBase;
	SCACCESSPOINTS : L_TS2P_scAP_SyncPosBase;
	MASTERVALUES : L_MC1P_IAXIS_REF_MASTERVALUES;
	XSYNCIN : BOOL;
	XSYNCPOSRESTORE : BOOL;
	LRSETBASEVEL : LREAL;
	LRSETOFFSETPOS : LREAL;
	XTRIMPOS : BOOL;
	XTRIMNEG : BOOL;
	XTRIMRESET : BOOL;
END_VAR
VAR_OUTPUT
	XREADYFOROPERATION : BOOL;
	XOPERATIONENABLED : BOOL;
	XREADYFORMOTION : BOOL;
	XERROR : BOOL;
	XWARNING : BOOL;
	EERRORID : L_IE1P_Error;
	XSTOACTIVE : BOOL;
	XQSPACTIVE : BOOL;
	XABORTBUSY : BOOL;
	XABORTDONE : BOOL;
	XJOGGINGBUSY : BOOL;
	XHOMINGBUSY : BOOL;
	XHOMINGDONE : BOOL;
	XISHOMED : BOOL;
	ETMSTATE : L_TB2P_States := L_TB2P_States.DISABLED;
	SCSTATUSBASICMOTION : L_TB2P_scStatusBasicMotion;
	LRACTVEL : LREAL;
	LRSETVELOUT : LREAL;
	LRACTPOS : LREAL;
	LRSETPOSOUT : LREAL;
	LRACTFOLLOWINGERROR : LREAL;
	SCSIGNALFLOW : L_TS2P_scSF_SyncPosBase;
	XSYNCHRONISED : BOOL;
	XACCDECSYNC : BOOL;
	XOFFSETTRIMACTIVE : BOOL;
	XBASEVELOCITYACTIVE : BOOL;
	LROFFSETTOTAL : LREAL;
END_VAR
VAR_IN_OUT
	AXIS : AXIS_REF;
END_VAR
VAR
	TM_INT : L_TS2P_TM_SyncPosBase_V2 := STRUCT(ModuleHandler := ModuleHandler);
	XENABLEOLD : BOOL;
END_VAR
END_FUNCTION_BLOCK

(* ---- L_TS2P_SYNCRONISEDOVERRIDE.fb ---- *)
FUNCTION_BLOCK L_TS2P_SYNCRONISEDOVERRIDE
VAR_INPUT
	XENABLE : BOOL;
	XSYNCHRONISED : BOOL;
	XEXECUTEGAP : BOOL;
	XAUXEXECUTEGAP : BOOL;
	LRSYNCOVERRIDE : LREAL := 1;
	LRCYCMASTERPOS : LREAL;
	LRCYCMASTERVEL : LREAL;
	LRCYCMASTERACC : LREAL;
	LRCYCSLAVEPOS : LREAL;
	LRCYCSLAVEVEL : LREAL;
	LRCYCSLAVEACC : LREAL;
	LRACC : LREAL;
	LRDEC : LREAL;
	LRJERK : LREAL;
	LRTASKCYLCETIME : LREAL := 0.001;
END_VAR
VAR_OUTPUT
	XBUSY : BOOL;
	XERROR : BOOL;
	EERRORID : L_IE1P_Error;
	XOVERRIDELIMITED : BOOL;
	XEXECUTEGAPOUT : BOOL;
	XAUXEXECUTEGAPOUT : BOOL;
	LRSETPOS : LREAL;
	LRSETVEL : LREAL;
	LRSETACC : LREAL;
	XSYNCOVERRIDEACTIVE : BOOL;
	XRAMPGENBUSY : BOOL;
END_VAR
VAR
	XENABLE_OLD : BOOL;
	XEXECUTEGAP_OLD : BOOL;
	XAUXEXECUTEGAP_OLD : BOOL;
	LRSYNCOVERRIDE_INT : LREAL := 1;
	LRSYNCOVERRIDE_LOCK : LREAL;
	LRADDOVERRIDE_LOCK : LREAL;
	WSTATE : WORD := 0;
	LROFFSETPOS_INT : LREAL;
	LROFFSETVEL_INT : LREAL;
	LROFFSETACC_INT : LREAL;
	LROFFSETVEL_OLD : LREAL;
	LRVELTARGET : LREAL;
	LRVELSTART : LREAL;
	FB_RAMPGENERATOR1 : L_MC1P_RampGenerator;
	C_LRCYCLELENGTHMASTER : LREAL := (16#4FFFFFFFFFFFFFFF * 1E-08);
END_VAR
END_FUNCTION_BLOCK

METHOD CALL_ERRORHANDLER
END_METHOD

METHOD CALL_FB_RAMPGENERATOR1
END_METHOD

METHOD CALL_OUTPUTS
END_METHOD

METHOD CALL_RESETCOMMANDS
END_METHOD

METHOD CALL_RESETOUTPUTS
END_METHOD

METHOD CALL_STATEMACHINE
END_METHOD

(* ---- L_TS2P_TM_CROSSCUTTERBASE.fb ---- *)
FUNCTION_BLOCK L_TS2P_TM_CROSSCUTTERBASE EXTENDS L_TB2P_SyncMotionControl
VAR_OUTPUT
	PAP : POINTER TO L_TS2P_scAP_TM_CrossCutterHigh;
	PSF : POINTER TO L_TS2P_scSF_TM_CrossCutterHigh;
	PPAR : POINTER TO L_TS2P_scPar_TM_CrossCutterHigh := ADR(scPar_int);
	PPARBASE : POINTER TO L_TS2P_scPar_TM_CrossCutterBaseExtension := ADR(scPar_int);
END_VAR
VAR_IN_OUT
	XEXECUTEMOVETOPARKPOS : BOOL;
	XSYNCIN : BOOL;
	XHOLDINPARKPOS : BOOL;
	LRPRODUCTLENGTH : LREAL;
	LROVERSPEED : LREAL;
	LRSETOFFSETPOSX : LREAL;
	XTRIMPOS : BOOL;
	XTRIMNEG : BOOL;
	XTRIMRESET : BOOL;
	SCSIGNALFLOW : L_TS2P_scSF_TM_CrossCutterBase;
	XSYNCHRONISED : BOOL;
	XACCDECSYNC : BOOL;
	XOFFSETTRIMACTIVE : BOOL;
	LROFFSETTOTAL : LREAL;
	XHOLDINPARKPOSACTIVE : BOOL;
	XCUTTINGACTIVE : BOOL;
	XCUTDONE : BOOL;
	LRACTCUTLENGTH : LREAL;
	XINPARKPOS : BOOL;
END_VAR
VAR
	TM_CROSSCUTTERBASECONFIG : L_TB2P_ModuleHandlerConfig;
	LROFFSET : LREAL;
	LROFFSETTRIM : LREAL;
	XEXECUTEMOVETOPARKPOS_INT : BOOL;
	XSYNCIN_INT : BOOL;
	XSYNCOUTINSTANT_INT : BOOL;
	XHOLDINPARKPOS_INT : BOOL;
	PMASTERAXIS : POINTER TO _AXIS_REF_REAL;
	LRPRODUCTLENGTH_INT : LREAL;
	LROVERSPEED_INT : LREAL;
	LRCUTTINGANGLE_INT : LREAL;
	LRSETOFFSETPOSX_INT : LREAL;
	LRSETOFFSETSLAVE_INT : LREAL;
	XTRIMPOS_INT : BOOL;
	XTRIMNEG_INT : BOOL;
	XRESETTRIMOFFSET_INT : BOOL;
	SCPAR_INT : L_TS2P_scPar_TM_CrossCutterHigh;
	SCPARBASE_INT : L_TS2P_scPar_TM_CrossCutterBaseExtension;
	LRSLAVEMAXVEL_INT : LREAL;
	LRSLAVEMAXACC_INT : LREAL;
	XCUTTINGBUSY_INT : BOOL;
	XACCDECSYNC_INT : BOOL;
	XCCMOVEABSEXECUTE_INT : BOOL;
	LRCCPOS_DIST_INT : LREAL;
	BYSETTOOLNOOUT : BYTE;
	BYSETAREAOUT : BYTE;
	LRSETXPOSOUT : LREAL;
	LRSETXVELOUT : LREAL;
	LRSETXACCOUT : LREAL;
	LRSLAVEMAXVEL : LREAL;
	LRSLAVEMAXACC : LREAL;
	LRMASTERVEL : LREAL;
	LRMASTERVEL_OLD : LREAL;
	LRMASTERVEL_OLD2 : LREAL;
	LRMASTERPOS_OLD : LREAL;
	LRACTMASTERPOS_OLD : LREAL;
	XMASTERAXISENABLED : BOOL;
	XMASTERAXISENABLED_OLD : BOOL;
	XCUTTINGACTIVE_OLD : BOOL;
	XRESETTRIMOFFSET_OLD : BOOL;
	XENABLECONTROLSETVALUES_OLD : BOOL;
	XINPARKPOS_OLD : BOOL;
	XMASTERISSTANDSTILL : BOOL;
	XNEXTTOOLDIRECTIONPOSITIV : BOOL := TRUE;
	ECUTTINGPROCESSSTATE : L_TB2P_States := L_TB2P_States.DISABLED;
	BYPOSITIONINGSTATE : BYTE := 0;
	BYMASTEROFFSETSTEPPER : BYTE := 0;
	BYTOOLCIRCARRAYPREPARED : BYTE;
	XMASTERIS_FREEENCODER : BOOL;
	XEXECUTETRANSITIONCYCLES : BOOL;
	XINVALIDCROSSCUTTERPARAMETRS : BOOL;
	XINVALIDCUTTINGPARAMETRS : BOOL;
	XMASTERNOTROTATIVE : BOOL;
	XWARNINGINVALIDPRODUCTLENGTH : BOOL;
	XINVALIDPRODUCTLENGTH : BOOL;
	XINVALIDCUTTINGANGLE : BOOL;
	XSLAVEOUTOFSCALE : BOOL;
	XERRORSLAVENOTINPARKPOS : BOOL;
	XMASTEROUTOFSCALE : BOOL;
	XSLAVERECEIVEDGAPS : BOOL;
	XINVALIDCAMSELECTED : BOOL;
	XWARNINGINVALIDCAMSELECTED : BOOL;
	XWARNINGDIRECTIONDISABLEDSYNCINT : BOOL;
	XWARNINGAXISNOTHOMED4SYNCIN : BOOL;
	ILOOPCNTR : INT;
	UIVARTEMP : UINT;
	IVARTEMP : INT;
	LRVARTEMP : LREAL;
	LRVARTEMP2 : LREAL;
	LRVARTEMP3 : LREAL;
	LRVARTEMP4 : LREAL;
	LRTEMPSTOPLENGTH : LREAL;
	LRTEMPSTARTLENGTH : LREAL;
	LRXDISTINPARKPOS : LREAL;
	XXPOSSYNCRONISEDMASTERPOS : BOOL;
	XCUTTINGPARISCHANGED : BOOL;
	XCAMDIRECTCHANGE_LOCK : BOOL;
	LRSETMASTERTRIMOFFSET_INT : LREAL;
	LRSETOFFSETMASTER_LOCK : LREAL;
	LRSETMASTERTRIMOFFSET_LOCK : LREAL;
	LRSETMASTERTRIMOFFSET_SAVE : LREAL;
	_LROFFSETTOTAL_OLD : LREAL;
	LRACTMASTERPOSSTART : LREAL;
	IMASTERPERIODCNT : INT;
	LRLENGTHCALCULATOR : LREAL;
	LROVERSPEEDUPPERLIMIT : LREAL := 2;
	ECUTTINGMODE_LOCK : L_TS2P_CuttingModeState;
	BYCAMCONTINUOUSNO_LOCK : BYTE := 1;
	BYNUMOFTOOLS_LOCK : BYTE;
	LRPRODUCTLENGTH_LOCK : LREAL;
	LRPRODUCTLENGTH_LOCK_OLD : LREAL;
	LRCUTLENGTH_LOCK : LREAL;
	LROSCILLATION_LOCK : LREAL := 0;
	LROVERSPEED_LOCK : LREAL;
	LROVERSPEEDFACTOR_LOCK : LREAL;
	LROVERSPEEDFACTOR_LOCK_OLD : LREAL;
	LRCUTTINGANGLE_LOCK : LREAL;
	LRSCALINGMASTER_LOCK : LREAL := 1;
	LRTOOLTOOLDIST_LOCK : LREAL;
	LRTOOLTOOLCIRCUMFERENCEDIST_LOCK : LREAL;
	LRCIRCUMFERENCE_LOCK : LREAL;
	LRCIRCUMFERENCEINV_LOCK : LREAL;
	XHOLDINPARKPOS_LOCK : BOOL;
	LRFACTOR_ANGLETOSLAVEUNITS_LOCK : LREAL;
	LRFACTOR_ANGLETOMASTERUNITS_LOCK : LREAL;
	LRFACTOR_SLAVEUNITSTOMASTERUNITS_LOCK : LREAL;
	LRFACTOR_MASTERUNITSTOSLAVEUNITS_LOCK : LREAL;
	LRFACTOR_PRODUCTUNITSTOMASTERUNITS_LOCK : LREAL;
	LRFACTOR_PRODUCTUNITSTOMASTERUNITSINV_LOCK : LREAL;
	LRFACTOR_PRODUCTUNITSTOMASTERUNITSINV_OLD : LREAL;
	XFIRSTCUT : BOOL;
	XCONTINUOUSMODE : BOOL := TRUE;
	BYSETCAMTABLENO : BYTE;
	BYREQUESTSSETCAMTABLE : BYTE;
	BYREQUESTSSETCAMTABLE_OLD : BYTE;
	SCSYNCSTARTLENGTH : L_MC2P_CamDataXYVA;
	SCSYNCSTOPLENGTH : L_MC2P_CamDataXYVA;
	SCASYNCLENGTH : L_MC2P_CamDataXYVA;
	SCSTARTLENGTH : L_MC2P_CamDataXYVA;
	SCSTOPLENGTH : L_MC2P_CamDataXYVA;
	LRSTANDSTILLLENGTH : LREAL;
	LRY_START : LREAL := 0;
	LRY_PARK : LREAL := 180;
	LRY_END : LREAL := 360;
	LRX_START : LREAL := 0;
	LRX_ENDSYNCPOS : LREAL := 10;
	LRX_STARTPARKPOS : LREAL := 180;
	LRX_ENDPARKPOS : LREAL := 180;
	LRX_STARTSYNCPOS : LREAL := 350;
	LRX_END : LREAL := 360;
	LRY_END_PREVIOUSLY : LREAL := 360;
	LRY_CUTLENGTHCALCULATOR : LREAL := 360;
	LROVERSPEED_LOCK_PREVIOUSLY : LREAL;
	FM_CAMCREATOR_START : L_TS2P_CamCreator;
	FM_CAMCREATOR_STOP : L_TS2P_CamCreator;
	FM_CAMCREATOR_CONTINUOUS : ARRAY [1..2] OF L_TS2P_CamCreator;
	FM_CAMCREATOR_STANDSTILL : L_TS2P_CamCreator;
	CAM_START_P : ARRAY [0..3] OF L_MC2P_CamDataXYVA;
	CAM_STOP_P : ARRAY [0..3] OF L_MC2P_CamDataXYVA;
	CAM_CONTINUOUS_P : ARRAY [1..2] OF ARRAY [0..3] OF L_MC2P_CamDataXYVA;
	CAM_STOPSTART_P : ARRAY [1..2] OF ARRAY [0..5] OF L_MC2P_CamDataXYVA;
	CAM_STANDSTILL_P : ARRAY [0..1] OF L_MC2P_CamDataXYVA;
	CAMTABLEATFLEXCAM : MC_CAM_REF;
	LRYOFFSET : LREAL;
	LRENDOFPROFILEWINDOWSIZE : LREAL := 0;
	_FC_XMASTERABSOLUTE : BOOL;
	_FC_XSLAVEABSOLUTE : BOOL;
	_FC_XPERIODIC : BOOL;
	_FC_XTRIMMASTERNEG : BOOL;
	_FC_XTRIMMASTERPOS : BOOL;
	_FC_LRSETOFFSETMASTER : LREAL;
	_FC_LRSETOFFSETSLAVE : LREAL;
	_FC_EPOSCTRLDIRECTION : L_MC2P.L_MC2P_ReverseCtrlDirection;
	_FC_EOFFSETMODEMASTER : L_MC2P.L_MC2P_OffsetMode;
	_FC_EOFFSETMODESLAVE : L_MC2P.L_MC2P_OffsetMode;
	_FC_XHOLDPROFGENMASTER : BOOL;
	_FC_ESYNCMODE : L_MC2P.L_MC2P_ClutchMode;
	_FC_ESYNCDIRECTION : L_MC2P.L_MC2P_ClutchDirection;
	_FC_LRMASTERSYNCINDIST : LREAL;
	_FC_LRMASTERSYNCINPOS : LREAL;
	_FC_LRMASTERSYNCOUTDIST : LREAL;
	_FC_LRSLAVESYNCOUTPOS : LREAL;
	_FC_LRSYNCINTIME : LREAL;
	_FC_LRSYNCOUTTIME : LREAL;
	_FC_LRSYNCOUTINSTANTDEC : LREAL;
	_FC_XENABLE : BOOL;
	_FC_XSYNCPOS : BOOL;
	_FC_XSYNCCAM : BOOL;
	_FC_XDIRECTCHANGE : BOOL;
	_FC_XSYNCOUTINSTANT : BOOL;
	_FC_LRSYNCCAMVEL : LREAL;
	_FC_LRSYNCCAMACC : LREAL;
	_FC_LRSYNCCAMDEC : LREAL;
	_FC_LRSYNCCAMJERK : LREAL;
	_FC_LRSETXPOSOUT : LREAL;
	_FC_LRSETXVELOUT : LREAL;
	_FC_LRSETXACCOUT : LREAL;
	_FC_LRSETYPOSOUT : LREAL;
	_FC_LRSETYVELOUT : LREAL;
	_FC_LRSETYACCOUT : LREAL;
	_FC_LRSETSLAVEPOSOUT : LREAL;
	_FC_LRSETSLAVEVELOUT : LREAL;
	_FC_LRSETSLAVEACCOUT : LREAL;
	_FC_XENDOFPROFILE : BOOL;
	_FC_XACCDECSYNC : BOOL;
	_FC_XSYNCHRONISED : BOOL;
	_FC_LRSETOFFSETMASTEROUT : LREAL;
	_FC_XENDOFCYCLE : BOOL;
	_FC_LRSETXPOS : LREAL;
	_FC_XCAMSYNCHRONISED : BOOL;
	_FC_XDONE : BOOL;
	_FC_XBUSY : BOOL;
	_FC_LRSETMASTERTRIMOFFSETOUT : LREAL;
	_FC_XENDOFPROFNEGATIVE : BOOL;
	_FC_LWENDOFPROFILECHECKSUM : LWORD;
	FM_FLEXCAMHIGH : L_MC2P_FlexCamHigh;
	FB_CONTROLSETVALUES : L_MC1P_ControlSetValues := STRUCT(eSetValueMode := L_MC1P_SetValueMode.Pos);
	L_MB1P_DIFFERENTIATE1 : L_MC2P_Differentiate;
	XINTERNALERROR : BOOL;
	WINTERNALERRORID : WORD;
	LWTCHECKSUM_INT : LWORD;
END_VAR
END_FUNCTION_BLOCK

METHOD CALL_ALLOCPOINTADR
END_METHOD

METHOD CALL_CTRLREQACTIVE : BOOL
END_METHOD

METHOD CALL_ERRORHANDLER
END_METHOD

METHOD CALL_ERRORHANDLER_STATECUTTING
END_METHOD

METHOD CALL_FBMETHODS
END_METHOD

METHOD CALL_FBMETHODS_BEFOREFLEXCAM
END_METHOD

METHOD CALL_FBMETHODS_CONTROLAXISBYPOS
END_METHOD

METHOD CALL_FB_CONTROLSETVALUES
END_METHOD

METHOD CALL_FB_DIFFERENTIATEPOSITION
END_METHOD

METHOD CALL_FM_CAMCREATOR_CONTINUOUS1
END_METHOD

METHOD CALL_FM_CAMCREATOR_CONTINUOUS2
END_METHOD

METHOD CALL_FM_CAMCREATOR_START
END_METHOD

METHOD CALL_FM_CAMCREATORS
END_METHOD

METHOD CALL_FM_FLEXCAM
END_METHOD

METHOD CALL_FM_FLEXCAM_INPUT
END_METHOD

METHOD CALL_INITDONE
END_METHOD

METHOD CALL_INITROUTINE
END_METHOD

METHOD CALL_INTERNALCTRL
END_METHOD

METHOD CALL_INTERNALCTRLBASEEXTENSION
END_METHOD

METHOD CALL_MASTEROFFSET
END_METHOD

METHOD CALL_MASTERTRIMM
END_METHOD

METHOD CALL_OUTPUT
END_METHOD

METHOD CALL_OUTPUTMINMAXVALUES
END_METHOD

METHOD CALL_OUTPUT_SF
END_METHOD

METHOD CALL_PARSYNCINCAM
END_METHOD

METHOD CALL_PARSYNCOUT
END_METHOD

METHOD CALL_REQUESTSSETCAMTABLE
END_METHOD

METHOD CALL_REQUESTSSETCAMTABLECTRL
END_METHOD

METHOD CALL_REQUESTS_EXT
END_METHOD

METHOD CALL_RESETCOMMANDS
END_METHOD

METHOD CALL_RESETOUTPUT
END_METHOD

METHOD CALL_RESETWARNINGS
END_METHOD

METHOD CALL_SETTOOLNOOUT
END_METHOD

METHOD CALL_STATEMACHINE
END_METHOD

METHOD CALL_ABC_INPUT
END_METHOD

METHOD CALL_ABC_INPUT_PROFILEPARAMETER
END_METHOD

METHOD CALL_CALCACTXKOORDINATEN
END_METHOD

METHOD CALL_CALCCAM_CONTINUOUS
END_METHOD

METHOD CALL_CALCCAM_START
END_METHOD

METHOD CALL_CALCSYNCARRAY
END_METHOD

METHOD CALL_CHECKCUTTINGPARCHANGES
END_METHOD

METHOD CALL_CONTINUOUSCAMSETYOFFSET
END_METHOD

METHOD CALL_CUTLENGTHCALCULATOR
END_METHOD

METHOD CALL_INIT_FLEXCAM
END_METHOD

METHOD CALL_LOCKCAMTABLE
END_METHOD

METHOD CALL_LOCKCROSSCUTTERPAR
END_METHOD

METHOD CALL_LOCKCUTTINGPAR
END_METHOD

METHOD CALL_LOCKCUTTINGPAR_ECCMODE_0
END_METHOD

METHOD CALL_LOCKCUTTINGPAR_ECCMODE_1
END_METHOD

METHOD CALL_PREPARENEXTCUT
END_METHOD

METHOD CALL_PREPARENEXTCUT_ECCMODEPAR
END_METHOD

METHOD CALL_RESETALLCAMCREATOR
END_METHOD

METHOD CALL_SEARCHACTYCOORDINATE
END_METHOD

METHOD CALL_SEARCHPARKPOS
END_METHOD

METHOD CALL_SETNEXTCAMCREATOR_CONTINUOUS
END_METHOD

METHOD CALL_YCOORDINATEMANAGER
END_METHOD

METHOD CHECKSLAVENOTINPARKPOS : BOOL
VAR_INPUT
	LRSETYPOS : LREAL;
	LRYSTART : LREAL;
	LRYPARK : LREAL;
	LRYEND : LREAL;
END_VAR
END_METHOD

METHOD CALL_CP_000_CYCLIC
END_METHOD

METHOD CALL_CP_001_INIT
END_METHOD

METHOD CALL_CP_001_INIT_OLD
END_METHOD

METHOD CALL_CP_141_IN_PARK_POS
END_METHOD

METHOD CALL_CP_142_ASYNC_PHASE
END_METHOD

METHOD CALL_CP_143_ENTRY_IN_SYNC_PHASE
END_METHOD

METHOD CALL_CP_143_ENTRY_IN_SYNC_PHASE_TRANSITION
END_METHOD

METHOD CALL_CP_144_EXIT_SYNC_PHASE
END_METHOD

METHOD CALL_CP_144_EXIT_SYNC_PHASE_TRANSITION
END_METHOD

METHOD CALL_CP_145_START_CAM
END_METHOD

METHOD CALL_CP_146_STOP_CAM
END_METHOD

METHOD CALL_CP_148_HOLD_IN_PARK_POS
END_METHOD

METHOD CALL_CP_148_HOLD_IN_PARK_POS_CONTINUECUTTING
END_METHOD

METHOD CALL_CP_148_HOLD_IN_PARK_POS_ENDOFPROFILE
END_METHOD

METHOD CALL_CP_802_STOP_IN_PARK_POS
END_METHOD

METHOD CALL_CP_900_DONE
END_METHOD

METHOD CALL_CUTTING_PROCESS
END_METHOD

METHOD CALL_S000_CYCLIC
END_METHOD

METHOD CALL_S002_STANDBY
END_METHOD

METHOD CALL_S030_SYNCHRONISING_POS
END_METHOD

METHOD CALL_S030_SYNCHRONISING_POS_ECCMODESELECT
END_METHOD

METHOD CALL_S030_SYNCHRONISING_POS_ECCMODE_0
END_METHOD

METHOD CALL_S030_SYNCHRONISING_POS_ECCMODE_1
END_METHOD

METHOD CALL_S032_POSITIONING_TO_START_POS
END_METHOD

METHOD CALL_S034_POSITIONING_TO_PARK_POS
END_METHOD

METHOD CALL_S035_CUTTING
END_METHOD

METHOD CALL_S996_STOP
END_METHOD

METHOD CALL_S999_ERROR
END_METHOD

METHOD CALL_T000_ALLSTATES
END_METHOD

METHOD CALL_S034_POSITIONING_TO_PARK_POS_OUT
END_METHOD

METHOD CALL_S035_CUTTING_OUT
END_METHOD

METHOD CALL_STATEMACHINE_OUT
END_METHOD

(* ---- L_TS2P_TM_CROSSCUTTERSTATE.fb ---- *)
FUNCTION_BLOCK L_TS2P_TM_CROSSCUTTERSTATE EXTENDS L_TS2P_TM_CrossCutterBase
VAR_IN_OUT
	SCTPRECDATA_MARKSENSOR : L_MC1P.L_MC1P_TpReceiveData;
	SCTPRECDATA_TOOLSENSOR : L_MC1P.L_MC1P_TpReceiveData;
	XTEACHMARKWINDOW : BOOL;
	XTEACHMARKWINDOWTOOL : BOOL;
	XGEARFACTORCORR : BOOL;
	XGEARFACTORCORRHOLD : BOOL;
	XTRQCTRLACTIVE : BOOL;
	LRSETMARKCORROUT : LREAL;
	XMARKWINDOWTEACHED : BOOL;
	LRGEARFACTORCORR : LREAL;
	LRSETTOOLCORROUT : LREAL;
	XMARKWINDOWTEACHEDTOOL : BOOL;
END_VAR
VAR
	XTEACHMARKWINDOW_INT : BOOL;
	XTEACHMARKWINDOWTOOL_INT : BOOL;
	XGEARFACTORCORR_INT : BOOL;
	XGEARFACTORCORRHOLD_INT : BOOL;
	LRCYCMASTERPOS_INT : LREAL;
	XLOADREGPOS_INT : BOOL;
	LRLOADREGPOS_INT : LREAL;
	LRSETMOTORPRECTRLTRQOUT : LREAL;
	XREGISTERCTRLACTIVE : BOOL;
	XMARKRECEIVED_OLD : BOOL;
	XTEACHMARKWINDOW_OLD : BOOL;
	XLOADREGPOS_OLD : BOOL;
	XMARKSENSORVALUESTORED_OLD : BOOL;
	AP11_XSETCUTLENGTHINPRODUCT_OLD : BOOL;
	EWARNINGID : WORD;
	FM_L_TS2P_MASTERVALUECORRECTION_LRACTVEL_OLD : LREAL;
	DNNUMAXISY_INT : DWORD := 1;
	DNDENAXISY_INT : DWORD := 1;
	XINVALIDCUTPRODUCTFORMAT : BOOL;
	XSCSCALINGVALID : BOOL := FALSE;
	XENABLETORQUEFOLLOWER : BOOL;
	XENABLEREGCTRLCORR : BOOL;
	XINVALIDTEACHMARKPOS : BOOL;
	XTPRECEIVED_INT : BOOL;
	LRTPACTPOSITION_INT : LREAL;
	XWARNINGINVALIDMARKRECIVED : BOOL;
	XTAKENEXTSTACKPOS : BOOL;
	LRSTACKLATESTDIST : LREAL;
	LRSENSORTOOLDIST_LOCK : LREAL;
	LRMARKPOS_LOCK : LREAL;
	XFIRSTCUTOFARRAY : BOOL;
	XCUTLENGTHINPRODUCTCHANGED_LOCK : BOOL;
	ISETNOCUTLENGTH_LOCK : INT;
	ISETNOOFMAXCUTLENGTH_LOCK : INT;
	LRUPPERCORRPOS_LOCK : LREAL;
	LRLOWERCORRPOS_LOCK : LREAL;
	ALRCUTLENGTHINPRODUCT_LOCK : ARRAY [1..10] OF LREAL;
	LRMARKSENSORPOS_LOCK : LREAL;
	LRREGISTERLENGTH_LOCK : LREAL;
	LRMINLOWERCORRPOS : LREAL;
	XCORRINSAMECYCLE : BOOL;
	LRFACTOR_NMOTOR_D_NAPPL : LREAL := 1;
	LRFACTOR_NAPPL_D_NMOTOR : LREAL := 1;
	LRFACTOR_MMOTOR_D_MAPPL : LREAL;
	INUMOFCUTLENGTH_LOCK : INT;
	INUMOFCUTLENGTH_INT : INT;
	LRREGPOS_ENDCUT : LREAL := 360;
	LRX_STOPCAMEND : LREAL := 360;
	_XSTACKENABLE : BOOL;
	_RC_LRUPPERCORRPOS : LREAL;
	_RC_LRLOWERCORRPOS : LREAL;
	_RC_XENABLE : BOOL;
	_RC_XMARKWINDOWOPEN : BOOL;
	_RC_XMARKOUTOFWINDOW : BOOL;
	_RC_XMARKNOTDETECTED : BOOL;
	_RC_XMARKWINDOWTEACHED : BOOL;
	_RC_LRGEARFACTORCORR : LREAL;
	_RC_XGEARFACTORCORRLIMITED : BOOL;
	_RC_LRPOSOUT : LREAL;
	_RC_LRACTVEL : LREAL;
	_RC_XERROR : BOOL;
	_RC_WERRORID : WORD;
	_RC_XLIMITACTIVE : BOOL;
	_RC_LRACTMARKERROR : LREAL;
	_RC_LRACTMARKDIST : LREAL;
	_RC_XINITDONE : BOOL;
	_RC_XCORRACTIVE : BOOL;
	_RC_XMARKRECEIVED : BOOL;
	_RC_LRREGMARKPOS : LREAL;
	_RC_XSETREGPOS2MASTERPOS : BOOL;
	LRACTMARKPOSDIFF : LREAL;
	FM_L_TS2P_MASTERVALUECORRECTION : L_TS2P_MasterValueCorrection;
	FM_L_TS2P_TOOLCORRECTION : L_TS2P_ToolCorrection;
	FB_L_TB2P_TP_CONVERTER : L_TB2P_TP_Converter;
	ITPCONVERTTPENABLECNTR : INT;
	FB_SETTORQUE1 : L_MC1P_SetTorqueOffset;
	FB_STACK : L_MB1P_Stack;
	WRESTART_LOCK : WORD;
	SCCAMTABLE_INT : MC_Cam_REF;
	SCSETXPROFILE_TEMP : L_MC2P_AxisProfile;
	SCSETYPROFILE_TEMP : L_MC2P_AxisProfile;
	PCAMDATA : POINTER TO L_MC2P_CamData;
	C_INUMOFCUTLENGTH : INT := 10;
END_VAR
END_FUNCTION_BLOCK

METHOD CALL_FM_TOOLCORRECTION : BOOL
END_METHOD

METHOD CALL_FM_TOOLCORRECTION_INPUT : BOOL
END_METHOD

METHOD CALL_ALLOCPOINTADRBASEEXTENSION
END_METHOD

METHOD CALL_ERRORHANDLER
END_METHOD

METHOD CALL_ERRORHANDLER_STATECUTTING
END_METHOD

METHOD CALL_FBMETHODS
END_METHOD

METHOD CALL_FBMETHODS_BEFOREFLEXCAM
END_METHOD

METHOD CALL_FBMETHODS_CONTROLAXISBYPOS
END_METHOD

METHOD CALL_FB_L_TB2P_TP_CONVERTER
END_METHOD

METHOD CALL_FB_SETTORQUE
END_METHOD

METHOD CALL_FB_SETTORQUE_INPUT
END_METHOD

METHOD CALL_FB_STACK
END_METHOD

METHOD CALL_FB_STACK_INPUT
END_METHOD

METHOD CALL_FM_CAMCREATOR_STANDSTILL
END_METHOD

METHOD CALL_FM_CAMCREATOR_STOP
END_METHOD

METHOD CALL_FM_CAMCREATORS
END_METHOD

METHOD CALL_FM_FLEXCAM
END_METHOD

METHOD CALL_FM_FLEXCAM_INPUT
END_METHOD

METHOD CALL_FM_REGISTERCONTROL
END_METHOD

METHOD CALL_FM_REGISTERCONTROL_INPUT
END_METHOD

METHOD CALL_FUN_GETSCALING
END_METHOD

METHOD CALL_INITDONE
END_METHOD

METHOD CALL_INITROUTINE
END_METHOD

METHOD CALL_INTERNALCTRL
END_METHOD

METHOD CALL_INTERNALCTRLBASEEXTENSION
END_METHOD

METHOD CALL_OUTPUT
END_METHOD

METHOD CALL_OUTPUTMINMAXVALUES
END_METHOD

METHOD CALL_OUTPUT_SF
END_METHOD

METHOD CALL_RESETCOMMANDS
END_METHOD

METHOD CALL_RESETOUTPUT
END_METHOD

METHOD CALL_RESETWARNINGS
END_METHOD

METHOD CALL_CALCCAM_RESTARTFROMSTOPCAM
END_METHOD

METHOD CALL_CALCCAM_STANDSTILL
END_METHOD

METHOD CALL_CALCCAM_STOP
END_METHOD

METHOD CALL_CALCSYNCARRAY_AP10STOPCAM
END_METHOD

METHOD CALL_CHECKARRAYOFCUTLENGTHCHANGES
END_METHOD

METHOD CALL_CHECKCUTPRODUCTFORMAT
END_METHOD

METHOD CALL_CHECKCUTTINGPARCHANGES
END_METHOD

METHOD CALL_CHECKRESTARTFROMSTOPCAM
END_METHOD

METHOD CALL_INIT_FLEXCAM
END_METHOD

METHOD CALL_LOCKCAMTABLE
END_METHOD

METHOD CALL_LOCKCROSSCUTTERPAR
END_METHOD

METHOD CALL_LOCKCUTTINGMODE
END_METHOD

METHOD CALL_LOCKCUTTINGPAR
END_METHOD

METHOD CALL_LOCKCUTTINGPAR_ECCMODE_2
END_METHOD

METHOD CALL_LOCKCUTTINGPAR_ECCMODE_3
END_METHOD

METHOD CALL_LOCKREGISTERCONTROLPAR
END_METHOD

METHOD CALL_PREAPAREARRAYOFCUTLENGTH
END_METHOD

METHOD CALL_PREPARENEXTCUT_ECCMODEPAR
END_METHOD

METHOD CALL_PREPARENEXTCUT_ECCMODEPAR_ECCMODE_2
END_METHOD

METHOD CALL_PREPARENEXTCUT_ECCMODEPAR_ECCMODE_3
END_METHOD

METHOD CALL_CP_000_CYCLIC
END_METHOD

METHOD CALL_CP_001_INIT
END_METHOD

METHOD CALL_CP_144_EXIT_SYNC_PHASE
END_METHOD

METHOD CALL_CP_148_HOLD_IN_PARK_POS
END_METHOD

METHOD CALL_CP_148_HOLD_IN_PARK_POS_CONTINUECUTTING
END_METHOD

METHOD CALL_CP_148_HOLD_IN_PARK_POS_ENDOFPROFILE
END_METHOD

METHOD CALL_CP_801_WAIT_OF_NEXT_CUT
END_METHOD

METHOD CALL_CP_802_STOP_IN_PARK_POS
END_METHOD

METHOD CALL_CP_900_DONE
END_METHOD

METHOD CALL_CUTTING_PROCESS
END_METHOD

METHOD CALL_S000_CYCLIC
END_METHOD

METHOD CALL_S002_READY
END_METHOD

METHOD CALL_S030_SYNCHRONISING_POS
END_METHOD

METHOD CALL_S030_SYNCHRONISING_POS_ECCMODESELECT
END_METHOD

METHOD CALL_S030_SYNCHRONISING_POS_ECCMODE_2
END_METHOD

METHOD CALL_S032_POSITIONING_TO_START_POS
END_METHOD

METHOD CALL_S999_ERROR
END_METHOD

(* ---- L_TS2P_TM_ELECTRONICGEARBOXBASE.fb ---- *)
FUNCTION_BLOCK L_TS2P_TM_ELECTRONICGEARBOXBASE EXTENDS L_TB2P_SyncMotionControl
VAR_OUTPUT
	PPAR : POINTER TO L_TS2P_scPar_TM_ElectronicGearboxBase := ADR(scPar_int);
	PSF : POINTER TO L_TS2P_scSF_TM_ElectronicGearboxBase;
	PAP : POINTER TO L_TS2P_scAP_TM_ElectronicGearboxBase;
END_VAR
VAR_IN_OUT
	XSYNCIN : BOOL;
	LRSETBASEVEL : LREAL;
	LRSETOFFSETPOS : LREAL;
	LRSETOFFSETVEL : LREAL;
	XTRIMPOS : BOOL;
	XTRIMNEG : BOOL;
	XTRIMRESET : BOOL;
	XINVERTGEARFACTOR : BOOL;
	SCSIGNALFLOW : L_TS2P_scSF_ElectronicGearboxBase;
	XSYNCHRONISED : BOOL;
	XACCDECSYNC : BOOL;
	XOFFSETTRIMACTIVE : BOOL;
	XBASEVELOCITYACTIVE : BOOL;
	LROFFSETTOTALVEL : LREAL;
END_VAR
VAR
	TM_ELECTRONICGEARBOXBASECONFIG : L_TB2P_ModuleHandlerConfig;
	LRSETBASEVEL_INT : LREAL := 0.0;
	XVELSYNCOUTTOBASESPEEDBUSY : BOOL;
	_LRSETBASEVEL : LREAL;
	XFM_SD_OFFSETBUSY : BOOL;
	_XSYNCHRONISEDBASEVEL : BOOL;
	XFM_SD_ACCDECBASEVEL : BOOL;
	_XSYNCOUTBASEVELDONE : BOOL;
	_XSYNCOUTBASEVELDONE_OLD : BOOL;
	_XSYNCOUTBASEVELDONE_RTRIG : BOOL;
	FM_L_TS2P_SYNCDRIVEVEL : L_TS2P_SyncDriveVel;
	XTRIMPOS_INT : BOOL;
	XTRIMNEG_INT : BOOL;
	XTRIMPOS_INT_OLD : BOOL;
	XTRIMNEG_INT_OLD : BOOL;
	XTRIMRESET_INT : BOOL;
	_XSYNCVEL : BOOL;
	_XSYNCOUTINSTANT : BOOL;
	_LRVELOFFSET : LREAL;
	_LRPOSOFFSETTOTALPOS : LREAL;
	_LRPOSOFFSETTOTALVEL : LREAL;
	_LROFFSETTOTALVEL : LREAL;
	_LRSETTRIMOFFSETOUT : LREAL;
	_XSYNCOUTDONE : BOOL;
	_XSYNCOUTDONE_OLD : BOOL;
	_XSYNCOUTDONE_RTRIG : BOOL;
	_XSYNCHRONISED : BOOL;
	_XACCDECSYNC : BOOL;
	_XOFFSETTRIMBUSY : BOOL;
	SCPAR_INT : L_TS2P_scPar_TM_ElectronicGearboxBase;
	XSYNCIN_INT : BOOL;
	LRSETOFFSETVEL_INT : LREAL;
	LRSETOFFSETPOS_INT : LREAL;
	XINVERTGEARFACTOR_INT : BOOL;
	DWGEARINGNUMERATOR_INT : DWORD;
	DWGEARINGDENOMINATOR_INT : DWORD;
	WMODE_INT : WORD;
	IACTMASTERDIRECTIONTMP : INT;
	XERROR_MODULOAXISISREQUIRED : BOOL;
	XERROR_INVALIDCOUPLINGMODE : BOOL;
	XWARNINGDIRECTIONDISABLEDSYNCINT : BOOL;
	XWARNINGDIRECTIONDISABLEDBASEVEL : BOOL;
	ETMSTATE_INT_TEMP : L_TB2P_States;
	XQSPAPPLICATION_OLD : BOOL;
	_XSYNCDRIVEENABLE : BOOL;
	_LRSYNCDRIVESETSLAVEVELOUT : LREAL;
	XENABLECONTROLSETVALUES : BOOL;
	FB_CONTROLSETVALUES : L_MC1P_ControlSetValues := STRUCT(eSetValueMode := L_MC1P_SetValueMode.VelAcc, xIgnoreAccForPosCalc := TRUE);
	FB_ALLOWEDDIRECTION : L_TS2P_AllowedDirection := STRUCT(eSetValueMode := L_MC1P_SetValueMode.VelAcc);
	XINVALIDBASEVELFLAG : BOOL;
	EERRORID_FIRST_OLD : L_IE1P_Error;
END_VAR
END_FUNCTION_BLOCK

METHOD CALL_FB_ALLOWEDDIRECTION
END_METHOD

METHOD CALL_ALLOCPOINTADR
END_METHOD

METHOD CALL_CTRLREQACTIVE : BOOL
END_METHOD

METHOD CALL_ERRORHANDLER
END_METHOD

METHOD CALL_FBMETHODS
END_METHOD

METHOD CALL_FB_CONTROLAXISBYVEL
END_METHOD

METHOD CALL_FB_CONTROLAXISBYVEL_INPUT
END_METHOD

METHOD CALL_FM_SYNCHRONIZEDDRIVE
END_METHOD

METHOD CALL_FM_SYNCHRONIZEDDRIVE_INPUT
END_METHOD

METHOD CALL_FM_SYNCHRONIZEDDRIVE_RESETFM
END_METHOD

METHOD CALL_INITDONE
END_METHOD

METHOD CALL_INITROUTINE
END_METHOD

METHOD CALL_INTERNALCTRL
END_METHOD

METHOD CALL_OUTPUT
END_METHOD

METHOD CALL_OUTPUT_SF
END_METHOD

METHOD CALL_REQUESTS_EXT
END_METHOD

METHOD CALL_RESETCOMMANDS
END_METHOD

METHOD CALL_RESETOUTPUT
END_METHOD

METHOD CALL_ABC
END_METHOD

METHOD CALL_ABC_INPUT_PROFILEPARAMETER
END_METHOD

METHOD CALL_S000_CYCLIC
END_METHOD

METHOD CALL_S001_INIT
END_METHOD

METHOD CALL_S002_STANDBY
END_METHOD

METHOD CALL_S003_HOMING
END_METHOD

METHOD CALL_S010_JOGGING
END_METHOD

METHOD CALL_S030_ACC_DEC_SYNC
END_METHOD

METHOD CALL_S031_SYNCHRONISED
END_METHOD

METHOD CALL_S051_BASEVELOCITY
END_METHOD

METHOD CALL_S996_STOP
END_METHOD

METHOD CALL_S999_ERROR
END_METHOD

METHOD CALL_STATEMACHINE
END_METHOD

METHOD CALL_T000_ALLSTATES
END_METHOD

METHOD CALL_T030_ACC_DEC_SYNC
END_METHOD

METHOD CALL_T031_SYNCHRONISED
END_METHOD

METHOD CALL_T051_BASEVELOCITY
END_METHOD

METHOD CALL_050_ABORT
END_METHOD

METHOD CALL_S000_CYCLIC_OUT
END_METHOD

METHOD CALL_S003_HOMING_OUT
END_METHOD

METHOD CALL_S010_JOGGING_OUT
END_METHOD

METHOD CALL_S014_MOVEABS_OUT
END_METHOD

METHOD CALL_S015_MOVEREL_OUT
END_METHOD

METHOD CALL_S996_STOP_OUT
END_METHOD

METHOD CALL_S999_ERROR_OUT
END_METHOD

METHOD CALL_STATEMACHINE_OUT
END_METHOD

METHOD CALL_T000_ALLSTATES_OUT
END_METHOD

(* ---- L_TS2P_TM_FLEXCAMBASE.fb ---- *)
FUNCTION_BLOCK L_TS2P_TM_FLEXCAMBASE EXTENDS L_TB2P_SyncMotionControl
VAR_OUTPUT
	PAP : POINTER TO L_TS2P_scAP_TM_FlexCamState;
	PPAR : POINTER TO L_TS2P_scPar_TM_FlexCamState := ADR(scPar_int);
	PSF : POINTER TO L_TS2P_scSF_TM_FlexCamState;
END_VAR
VAR_IN_OUT
	XSYNCIN : BOOL;
	XCAMCHANGEINSTANT : BOOL;
	LRSETOFFSETMASTER : LREAL;
	LRSETOFFSETSLAVE : LREAL;
	LRSETSCALINGMASTER : LREAL;
	LRSETSCALINGSLAVE : LREAL;
	CAMTABLE1 : MC_CAM_REF;
	SCSIGNALFLOW : L_TS2P_scSF_TM_FlexCamState;
	XCAMMINGBUSY : BOOL;
	XSYNCHRONISED : BOOL;
	XACCDECSYNC : BOOL;
	XENDOFPROFILE : BOOL;
	LROFFSETMASTER : LREAL;
	LROFFSETSLAVE : LREAL;
END_VAR
VAR
	TM_FLEXCAMBASECONFIG : L_TB2P_ModuleHandlerConfig;
	XSYNCIN_INT : BOOL;
	XSYNCOUTINSTANT_INT : BOOL;
	XCAMCHANGEINSTANT_INT : BOOL;
	LRSETOFFSETMASTER_INT : LREAL;
	LRSETOFFSETSLAVE_INT : LREAL;
	LRSETSCALINGMASTER_INT : LREAL := 1;
	LRSETSCALINGSLAVE_INT : LREAL := 1;
	SCPAR_INT : L_TS2P_scPar_TM_FlexCamState;
	XCAMMINGBUSY_INT : BOOL;
	XENABLECAMPROFILERSTANDBY_INT : BOOL := TRUE;
	XINTERNALCAMBASICACTIVE_INT : BOOL;
	XCAMCHANGEINSTANT_OLD : BOOL;
	LRMASTERVEL_OLD : LREAL;
	LRMASTERVEL_OLD2 : LREAL;
	LRMASTERPOS_OLD : LREAL;
	XCONTROLSETVALUESBUSY_OLD : BOOL;
	XMASTERABSOLUTE_OLD : BOOL;
	XCAMTABLEVALID_INT : BOOL;
	XERROR_INVALIDSYNCMODE : BOOL;
	XERROR_INVALIDCAMTABLE : BOOL;
	XWARNING_INVALIDCAMTABLE : BOOL;
	LRTRACEACCMAX_INT : LREAL;
	XCOMMUNICATION : BOOL;
	CAMTABLE_INIT : MC_CAM_REF;
	XMASTERPARCHANGED : BOOL;
	MASTERID : POINTER TO WORD;
	LRCYCLELENGTH : LREAL;
	ETRAVERSINGRANGE : LREAL;
	LRACTYPOS : LREAL;
	LRACTYVEL : LREAL;
	LRCAMYSTART : LREAL;
	LRCAMYEND : LREAL;
	LRACTIVESCALINGSLAVEINVERSE : LREAL;
	XCAMTABLEINTERNALVALID : BOOL;
	CAMTABLEINTERNAL : MC_CAM_REF;
	PCAMDATA : POINTER TO L_MC2P_CamData;
	_WFC_ENABLEMODE : WORD;
	_WFC_ENABLEMODE_OLD : WORD;
	_LRFC_SETXPOSOUT : LREAL;
	_LRFC_SETXVELOUT : LREAL;
	_LRFC_SETXACCOUT : LREAL;
	_LRFC_SETYPOSOUT : LREAL;
	_LRFC_SETYVELOUT : LREAL;
	_LRFC_SETYACCOUT : LREAL;
	_LRFC_OFFSETMASTER : LREAL;
	_LRFC_OFFSETSLAVE : LREAL;
	_XFC_CRITICALCYCLE : BOOL;
	_XFC_ENDOFPROFILE : BOOL;
	_XFC_ACCDECSYNC : BOOL;
	_XFC_CAMSYNCHRONISED : BOOL;
	_XFC_BUSY : BOOL;
	_XFC_DONE : BOOL;
	_XFC_ERROR : BOOL;
	_LRFC_SETSLAVEPOSOUT : LREAL;
	_LRFC_SETSLAVEVELOUT : LREAL;
	_LRFC_SETSLAVEACCOUT : LREAL;
	LRENDOFPROFILEWINDOWSIZE : LREAL := 0;
	MP_LRCONVERTMASTERTOXPOS : LREAL;
	MP_LRCAMPROFILERPOSOUT : LREAL;
	MP_LRCONVERTYTOSLAVEPOS : LREAL;
	MP_LWENDOFPROFILECHECKSUM : LWORD;
	MP_XENDOFPROFPOSITIVE : BOOL;
	MP_XENDOFPROFNEGATIVE : BOOL;
	SCSETXPROFILE : L_MC2P_AxisProfile;
	SCSETYPROFILE : L_MC2P_AxisProfile;
	FB_CAMBASIC : L_MC2P_CamBasic;
	FB_CONTROLSETVALUES : L_MC1P_ControlSetValues;
	FB_CAMTABLEINFO1 : L_TS2P_CamTableInfo;
END_VAR
END_FUNCTION_BLOCK

METHOD CALL_ALLOCPOINTADR
END_METHOD

METHOD CALL_AXISCONTROLBYPOS
END_METHOD

METHOD CALL_AXISCONTROLBYPOS_INPUT
END_METHOD

METHOD CALL_CAMBOUNDS
END_METHOD

METHOD CALL_CTRLREQACTIVE : BOOL
END_METHOD

METHOD CALL_CURVESKETCHING
END_METHOD

METHOD CALL_ERRORHANDLER
END_METHOD

METHOD CALL_FBMETHODS
END_METHOD

METHOD CALL_FB_CAMBASIC
END_METHOD

METHOD CALL_FM_CAMTABLEINFO1
END_METHOD

METHOD CALL_FM_FLEXCAM
END_METHOD

METHOD CALL_FM_FLEXCAM_INPUT
END_METHOD

METHOD CALL_INITDONE
END_METHOD

METHOD CALL_INITROUTINE
END_METHOD

METHOD CALL_INTERNALCTRL
END_METHOD

METHOD CALL_MASTERAXISREF
VAR_INPUT
	MASTERVALUES : L_MC1P_IAXIS_REF_MASTERVALUES;
END_VAR
END_METHOD

METHOD CALL_OUTPUT
END_METHOD

METHOD CALL_OUTPUTMINMAXVALUES
END_METHOD

METHOD CALL_OUTPUTMINMAXVALUESMODULOOVERRUN
END_METHOD

METHOD CALL_OUTPUTMINMAXVALUESOFCAMTABLES1
END_METHOD

METHOD CALL_OUTPUT_SF
END_METHOD

METHOD CALL_REQUESTS_EXT
END_METHOD

METHOD CALL_RESETCOMMANDS
END_METHOD

METHOD CALL_RESETOUTPUT
END_METHOD

METHOD CALL_STATEMACHINE
END_METHOD

METHOD CALL_ABC_INPUT
END_METHOD

METHOD CALL_ABC_INPUT_PROFILEPARAMETER
END_METHOD

METHOD CAMREFCHANGED : BOOL
VAR_IN_OUT
	CAMREFNEW : MC_CAM_REF;
	CAMREFOLD : MC_CAM_REF;
END_VAR
END_METHOD

METHOD CAMREFVALID : BOOL
VAR_INPUT
	CAMREF : MC_CAM_REF;
END_VAR
END_METHOD

METHOD GET_INTERNCAMTABLE : MC_CAM_REF
END_METHOD

METHOD GET_ECAMTYPE : L_MC2P_CamType
END_METHOD

METHOD GET_LRACTIVESCALINGSLAVE : LREAL
END_METHOD

METHOD GET_LRCAMXEND : LREAL
END_METHOD

METHOD GET_LRCAMXSTART : LREAL
END_METHOD

METHOD GET_LRCAMYEND : LREAL
END_METHOD

METHOD GET_LRCAMYSTART : LREAL
END_METHOD

METHOD GET_XCOMMUNICATION : BOOL
END_METHOD

METHOD RESET_SYSTEMFAULT
END_METHOD

METHOD SET_SYSTEMFAULT
VAR_INPUT
	IN : L_IE1P_Error;
END_VAR
END_METHOD

METHOD SET_ESTATE
VAR_INPUT
	IN : L_TB2P_States;
END_VAR
END_METHOD

METHOD CALL_S000_CYCLIC
END_METHOD

METHOD CALL_S002_STANDBY
END_METHOD

METHOD CALL_S112_CAMMING
END_METHOD

METHOD CALL_S112_CAMMING_RESTARTFLEXCAM
END_METHOD

METHOD CALL_S996_STOP
END_METHOD

METHOD CALL_S999_ERROR
END_METHOD

METHOD CALL_T000_ALLSTATES
END_METHOD

METHOD CALL_T002_STANDBY
END_METHOD

(* ---- L_TS2P_TM_FLEXCAMSTATE.fb ---- *)
FUNCTION_BLOCK L_TS2P_TM_FLEXCAMSTATE EXTENDS L_TS2P_TM_FlexCamBase
VAR_IN_OUT
	CAMTABLE2 : MC_CAM_REF;
	CAMTABLE3 : MC_CAM_REF;
	CAMTABLE4 : MC_CAM_REF;
	WSETCAMTABLE : WORD;
	XCAMSEQUENCER : BOOL;
	WACTIVECAMTABLE : WORD;
	XCAMSEQUENCERACTIVE : BOOL;
END_VAR
VAR
	WSETCAMTABLE_INT : WORD := 1;
	XCAMSEQUENCER_INT : BOOL;
	XSLAVEABSOLUTE_OLD : BOOL;
	XUPDATECURVE : BOOL;
	_XMCS_ENABLE : BOOL;
	_MCS_CAMTABLEOUT : MC_CAM_REF;
	FM_FLEXCAMSTATE1 : L_MC2P_FlexCamHigh := STRUCT(ePosCtrlDirection := L_MC2P_ReverseCtrlDirection.both);
	FB_MULTICAMSEQUENCER1 : L_TS2P_MultiCamSequencer;
	FB_CAMTABLEINFO2 : L_TS2P_CamTableInfo;
	FB_CAMTABLEINFO3 : L_TS2P_CamTableInfo;
	FB_CAMTABLEINFO4 : L_TS2P_CamTableInfo;
END_VAR
END_FUNCTION_BLOCK

METHOD CALL_CURVESKETCHING
END_METHOD

METHOD CALL_ERRORHANDLER
END_METHOD

METHOD CALL_FBMETHODS
END_METHOD

METHOD CALL_FM_CAMTABLEINFO2
END_METHOD

METHOD CALL_FM_CAMTABLEINFO3
END_METHOD

METHOD CALL_FM_CAMTABLEINFO4
END_METHOD

METHOD CALL_FM_FLEXCAM
END_METHOD

METHOD CALL_FM_FLEXCAM_INPUT
END_METHOD

METHOD CALL_FM_MULTICAMSEQUENCER
END_METHOD

METHOD CALL_FM_MULTICAMSEQUENCER_INPUT
END_METHOD

METHOD CALL_FIRSTCYCLE
END_METHOD

METHOD CALL_INTERNALCTRL
END_METHOD

METHOD CALL_OUTPUT
END_METHOD

METHOD CALL_OUTPUTMINMAXVALUES
END_METHOD

METHOD CALL_OUTPUTMINMAXVALUESOFCAMTABLES1
END_METHOD

METHOD CALL_OUTPUTMINMAXVALUESOFCAMTABLES1_2_3_4
END_METHOD

METHOD CALL_OUTPUT_SF
END_METHOD

METHOD CALL_RESETCOMMANDS
END_METHOD

METHOD CALL_RESETCOMMANDSFLEXCAM
END_METHOD

METHOD CALL_RESETOUTPUT
END_METHOD

METHOD FUN_FMSYNCDIRCTION : L_MC2P_ClutchMode
VAR_INPUT
	ESYNCMODE : L_TS2P_SyncModeFlexCam;
END_VAR
END_METHOD

METHOD GET_INTERNCAMTABLE : MC_CAM_REF
END_METHOD

METHOD GET_LRACTIVESCALINGSLAVE : LREAL
END_METHOD

METHOD GET_LRCAMXEND : LREAL
END_METHOD

METHOD GET_LRCAMXSTART : LREAL
END_METHOD

METHOD GET_LRCAMYEND : LREAL
END_METHOD

METHOD GET_LRCAMYSTART : LREAL
END_METHOD

METHOD CALL_S112_CAMMING_RESTARTFLEXCAM
END_METHOD

(* ---- L_TS2P_TM_FLYINGSAWSTATE_V2.fb ---- *)
FUNCTION_BLOCK L_TS2P_TM_FLYINGSAWSTATE_V2 EXTENDS L_TB2P_SyncMotionControl
VAR_OUTPUT
	PPAR : POINTER TO L_TS2P_scPar_TM_FlyingSawState := ADR(scPar_int);
	PSF : POINTER TO L_TS2P_scSF_TM_FlyingSawState;
	PAP : POINTER TO L_TS2P_scAP_TM_FlyingSawState;
END_VAR
VAR_IN_OUT
	XSTARTFLYINGSAW : BOOL;
	XSYNCININSTANT : BOOL;
	XEXECUTENEXTCUT : BOOL;
	XEXECUTEGAP : BOOL;
	XSETCUTTINGLENGTHINSTANT : BOOL;
	LRCUTTINGLENGTH : LREAL;
	XSETMATERIALCOUNTER : BOOL;
	LRSYNCOVERRIDE : LREAL;
	SCSIGNALFLOW : L_TS2P_scSF_FlyingSawState;
	XSYNCHRONISED : BOOL;
	XACCDECSYNC : BOOL;
	XPOSITIONING : BOOL;
	XINPOSITION : BOOL;
	LRMATERIALCOUNTER : LREAL;
	LRTARGETPOS : LREAL;
	LRCUTGAP : LREAL;
	LRACTIVECUTTINGLENGTH : LREAL;
	XMOVETOPARKPOS : BOOL;
	XRESUMETARGETPOS : BOOL;
	XRESETMARKSTACK : BOOL;
	SCTPRECDATA_MARKSENSOR : L_MC1P.L_MC1P_TpReceiveData;
	WMARKSINSTACK : WORD;
END_VAR
VAR
	TM_FLYINGSAWSTATECONFIG : L_TB2P_ModuleHandlerConfig;
	SCPAR_INT : L_TS2P_scPar_TM_FlyingSawState;
	XSTARTFLYINGSAW_INT : BOOL;
	XSYNCININSTANT_INT : BOOL;
	LRSETOFFSETSLAVE_INT : LREAL;
	XSETMATERIALCOUNTER_INT : BOOL;
	XEXECUTENEXTCUT_INT : BOOL;
	LRSYNCOVERRIDE_INT : LREAL := 1;
	XENABLEHWLIMIT_INT : BOOL;
	XHWLIMITPOS_INT : BOOL;
	XHWLIMITNEG_INT : BOOL;
	XEXECUTEGAP_INT : BOOL;
	XSETCUTTINGLENGTHINSTANT_INT : BOOL;
	LRCUTLENGTHPROCESSED : LREAL;
	LRDISTTOCUTPOSITION : LREAL;
	XACCDECSYNC_INT : BOOL;
	LROFFSET_STORE : LREAL;
	FB_MATERIALCOUNTER : L_TS2P_MaterialCounter;
	FB_CALCULATETARGETPOS : L_TS2P_CalculateTargetPos;
	FB_PROCESSCONTROL : L_TS2P_ProcessControl;
	FB_POSPROFILERCLUTCH : L_MB1P_PosProfilerClutchHigh;
	FB_CONTROLSETVALUES : L_MC1P_ControlSetValues;
	FB_L_TB2P_TP_CONVERTER : L_TB2P_TP_Converter;
	FB_STACK : L_MB1P_Stack;
	FB_SYNCRONISEDOVERRIDE : L_TS2P_SyncronisedOverride;
	RS_SYNCHRONISED : RS;
	WSTEPPER : wStepperFS;
	LRSTARTPOSOUT : LREAL;
	LRSTARTPOSOUT2 : LREAL;
	LRACCDIST : LREAL;
	LRACCTIME : LREAL;
	LRDECDIST : LREAL;
	LRDECTIME : LREAL;
	LRMASTERPOS1 : LREAL;
	LRMASTERPOS2 : LREAL;
	LRSLAVEPOS1 : LREAL;
	LRSLAVEPOS2 : LREAL;
	XSYNCHRONIZEDOLD : BOOL;
	WSTEPPER1 : WORD;
	LRCUTGAP_INT : LREAL;
	XGAPDONE : BOOL;
	WSTEPPER2 : WORD;
	LRCUTTINGLENGTH_INT : LREAL;
	LRDIST_INT : LREAL;
	XTIMESYNCINVALID : BOOL;
	LRTIMESYNCIN_INT : LREAL;
	EFLYINGSAWMODE_INT : L_TS2P_FlyingSawMode := L_TS2P_FlyingSawMode.MarkControlled;
	XRESETMARKSTACK_INT : BOOL;
	XTEST : BOOL;
	XTPRECEIVED_INT : BOOL;
	LRTPACTPOSITION_INT : LREAL;
	FB_INPOSITION : L_TT1P_InPosition;
	XMOVETOPARKPOS_INT : BOOL;
	XRESUMETARGETPOS_INT : BOOL;
	LRSYNCOUTPOS : LREAL;
	XNEXTCUT_IP : BOOL;
	WSTEPPERSKPCUT : INT;
	XSYNCINSTANT_IP : BOOL;
	XFIRSTTP : BOOL;
	XMODECHANGE : BOOL;
	XMODECHANGE_OLD : BOOL;
	XFIRSTTP_OLD : BOOL;
	EFLYINGSAWMODE_OLD : L_TS2P_FlyingSawMode;
	PAXISREAL : POINTER TO _AXIS_REF_REAL;
	BYTEST : BYTE;
	LRRANGEOFTOLERANCE : LREAL;
	XBALANCEDPROFILEACTIVE : BOOL;
	LRDISTTOTARGET : LREAL;
	LRFILTMATERIALVEL : LREAL;
	LRFILTMATERIALACC : LREAL;
	XMATERIALCONSTANTVEL : BOOL;
	LRRESTTIMETARGETTOLOWERLIMIT : LREAL;
	LRSETRESTTIMETARGETTOLOWERLIMIT : LREAL;
	_LRREGISTERCNTRFACTOR : LREAL;
	_LRTPAXISDELAYCYCLE : LREAL;
	_LRTPDELAYCYCLESACTPOS : LREAL;
	_DWTPAXISDELAYCYCLE : DWORD;
	_LRRESIDUAL : LREAL;
	XTACKEPOSINSTACK_INT : BOOL;
	XWARNING_TPRECPOSITIONNOTSUPPORTED : BOOL;
	XQSPAPPLICATION_OLD : BOOL;
	FB_STACKCONTROLARRAYNOISE : L_MC1P_StackControlArray := STRUCT(iMaxLegth := 10);
	ALRDELTAVEL : ARRAY [0..10] OF LREAL;
	AXNOISE : ARRAY [0..5] OF BOOL;
	ALRVELTOLERANCE : ARRAY [0..5] OF LREAL;
	XNOISE : BOOL;
	XACCPOSITIV : BOOL;
	IACCCHANGEDIRECTIONCOUNTER : INT;
	LRVELTOLERANCE_INT : LREAL;
	LRMAXVELTOLERANCE : LREAL;
	LRMAXACCTOLERANCE : LREAL;
	LRCYCMASTERVEL : LREAL;
	LRCYCMASTERVEL_OLD : LREAL;
	XEXECUTEMOVETOPARKPOS : BOOL;
	WABCMOVETOPARKPOSSTEPPER : WORD;
	LRPARKPOS : LREAL;
	XTMHALT_INT : BOOL;
	XTMHALT_OLD : BOOL;
	C_LRMATERIALCOUNTERCYCLELENGTH : LREAL := (16#4FFFFFFFFFFFFFFF * 1E-08);
END_VAR
END_FUNCTION_BLOCK

METHOD CALL_ALLOCPOINTADR
END_METHOD

METHOD CALL_CALCULATECUTTINGLENGTH
END_METHOD

METHOD CALL_CHECKMASTERNOISE : BOOL
END_METHOD

METHOD CALL_CTRLREQACTIVE : BOOL
END_METHOD

METHOD CALL_ERRORRESETACTIVE
END_METHOD

METHOD CALL_ERRORHANDLER
END_METHOD

METHOD CALL_FBMETHODS
END_METHOD

METHOD CALL_INITDONE
END_METHOD

METHOD CALL_INITROUTINE
END_METHOD

METHOD CALL_INTERNALCTRL
END_METHOD

METHOD CALL_OUTPUT
END_METHOD

METHOD CALL_OUTPUT_SF
END_METHOD

METHOD CALL_REQUESTS_EXT
END_METHOD

METHOD CALL_RESETCOMMANDS
END_METHOD

METHOD CALL_RESETOUTPUT
END_METHOD

METHOD CALL_STATEMACHINE
END_METHOD

METHOD CALL_ABC_INPUT
END_METHOD

METHOD CALL_ABC_INPUT_PROFILEPARAMETER
END_METHOD

METHOD CALL_FB_CALCULATETARGETPOS
END_METHOD

METHOD CALL_FB_CALCULATETARGETPOSINPUTS
END_METHOD

METHOD CALL_FB_CONTROLSETVALUES
END_METHOD

METHOD CALL_FB_CONTROLSETVALUESINPUTS
END_METHOD

METHOD CALL_FB_INPOSITION
END_METHOD

METHOD CALL_FB_INPOSITIONINPUTS
END_METHOD

METHOD CALL_FB_L_TB2P_TP_CONVERTER
END_METHOD

METHOD CALL_FB_MATERIALCOUNTER
END_METHOD

METHOD CALL_FB_MATERIALCOUNTERINPUTS
END_METHOD

METHOD CALL_FB_POSPROFILERCLUTCH
END_METHOD

METHOD CALL_FB_POSPROFILERCLUTCHINPUTS
END_METHOD

METHOD CALL_FB_PROCESSCONTROL
END_METHOD

METHOD CALL_FB_PROCESSCONTROLINPUTS
END_METHOD

METHOD CALL_FB_STACK
END_METHOD

METHOD CALL_FB_STACK_INPUTS
END_METHOD

METHOD CALL_FB_SYNCRONISEDOVERRIDE
END_METHOD

METHOD CALL_S000_CYCLIC
END_METHOD

METHOD CALL_S002_STANDBY
END_METHOD

METHOD CALL_S003_HOMING
END_METHOD

METHOD CALL_S010_JOGGING
END_METHOD

METHOD CALL_S030_SAW_IN_PROCESS
END_METHOD

METHOD CALL_S040_MOVE_TO_PARKPOS
END_METHOD

METHOD CALL_S996_STOP
END_METHOD

METHOD CALL_S999_ERROR
END_METHOD

METHOD CALL_T000_ALLSTATES
END_METHOD

METHOD CALL_T030_SAW_IN_PROCESS
END_METHOD

METHOD CALL_S000_CYCLIC_OUT
END_METHOD

METHOD CALL_S003_HOMING_OUT
END_METHOD

METHOD CALL_S010_JOGGING_OUT
END_METHOD

METHOD CALL_S013_MOVEVEL_OUT
END_METHOD

METHOD CALL_S014_MOVEABS_OUT
END_METHOD

METHOD CALL_S015_MOVEREL_OUT
END_METHOD

METHOD CALL_S017_EXTERNAL_OUT
END_METHOD

METHOD CALL_S996_STOP_OUT
END_METHOD

METHOD CALL_S999_ERROR_OUT
END_METHOD

METHOD CALL_STATEMACHINE_OUT
END_METHOD

METHOD CALL_T000_ALLSTATES_OUT
END_METHOD

METHOD CALL_S000_STARTSAW
END_METHOD

METHOD CALL_S020_SAWSYNCHRONIZED
END_METHOD

METHOD CALL_S030_MOVETOLOWERLIMIT
END_METHOD

METHOD CALL_S040_WAITINGFORNEXTCUT
END_METHOD

(* ---- L_TS2P_TM_SYNCANDCORRECTIONSTATE.fb ---- *)
FUNCTION_BLOCK L_TS2P_TM_SYNCANDCORRECTIONSTATE EXTENDS L_TS2P_TM_SyncPosBase
VAR_INPUT
	SCTPRECDATA_MARKSENSOR : L_MC1P.L_MC1P_TpReceiveData;
	SCTPRECDATA_TOOLSENSOR : L_MC1P.L_MC1P_TpReceiveData;
	XTEACHMARKWINDOW : BOOL;
	XTEACHMARKWINDOWTOOL : BOOL;
	XGEARFACTORCORR : BOOL;
	XGEARFACTORCORRHOLD : BOOL;
END_VAR
VAR_OUTPUT
	LRSETMARKCORROUT : LREAL;
	XMARKWINDOWTEACHED : BOOL;
	LRGEARFACTORCORR : LREAL;
	LRSETTOOLCORROUT : LREAL;
	XMARKWINDOWTEACHEDTOOL : BOOL;
END_VAR
VAR
	TM_SYNCANDCORRECTIONSTATECONFIG : L_TB2P_ModuleHandlerConfig;
	ITFSYNCANDCORRECTIONSTATE : L_TS2P_ISyncAndCorrectionState := THIS^;
	SCDATA_INTSC : L_TS2P_scData_TM_SyncAndCorrectionState;
	PAP_SC : POINTER TO L_TS2P_scAP_TM_SyncAndCorrectionState;
	PSF_SC : POINTER TO L_TS2P_scSF_TM_SyncAndCorrectionState;
	PDATASC : POINTER TO L_TS2P_scData_TM_SyncAndCorrectionState := ADR(scData_IntSC);
	PPAR_SC : POINTER TO L_TS2P_scPar_TM_SyncAndCorrectionState;
	FM_L_TS2P_MASTERVALUECORRECTION : L_TS2P_MasterValueCorrection;
	FM_L_TS2P_TOOLCORRECTION : L_TS2P_ToolCorrection;
	CONNECTOR : __SYSTEM.IQueryInterface;
	SYNCANDCORRECTIONSTATEEXTENSION : L_TS2P_ISyncAndCorrectionState;
	SYNCPOSBASEEXTENSION : L_TS2P_ISyncPosBase;
END_VAR
END_FUNCTION_BLOCK

METHOD CALLFBS
VAR_INPUT
	ECASE : L_UBUP_StateHandleCase;
END_VAR
END_METHOD

METHOD FINALIZECYCLE
END_METHOD

METHOD PREPARECYCLE
END_METHOD

METHOD SETADDMODULEINFO
VAR_INPUT
	ESUBCOMPTYPE : UDINT;
	SLICINFO : STRING(10);
END_VAR
END_METHOD

METHOD CALL_SETLOCALMASTERVALUES
END_METHOD

METHOD STATE_11_SYNC_ACC
VAR_INPUT
	ECASE : L_UBUP_StateHandleCase;
	ISTATESERVER : L_UBUP_IStateServer;
END_VAR
END_METHOD

METHOD CALL_FM_MASTERVALUECORRECTION
END_METHOD

METHOD CALL_FM_MASTERVALUECORRECTION_INPUT
END_METHOD

METHOD CALL_FM_TOOLCORRECTION : BOOL
END_METHOD

METHOD CALL_FM_TOOLCORRECTION_INPUT : BOOL
END_METHOD

METHOD CALL_ALLOCPOINTADR
END_METHOD

METHOD CALL_EXIT_CALLFBS
END_METHOD

METHOD CALL_INIT_CALLFBS
END_METHOD

METHOD CALL_INTERNALCTRL
END_METHOD

METHOD CALL_RESETOUTPUT
END_METHOD

(* ---- L_TS2P_TM_SYNCANDCORRECTIONSTATE_V2.fb ---- *)
FUNCTION_BLOCK L_TS2P_TM_SYNCANDCORRECTIONSTATE_V2 EXTENDS L_TS2P_TM_SyncPosBase_V2
VAR_IN_OUT
	SCTPRECDATA_MARKSENSOR : L_MC1P.L_MC1P_TpReceiveData;
	SCTPRECDATA_TOOLSENSOR : L_MC1P.L_MC1P_TpReceiveData;
	XTEACHMARKWINDOW : BOOL;
	XTEACHMARKWINDOWTOOL : BOOL;
	XGEARFACTORCORR : BOOL;
	XGEARFACTORCORRHOLD : BOOL;
	LRSETMARKCORROUT : LREAL;
	XMARKWINDOWTEACHED : BOOL;
	LRGEARFACTORCORR : LREAL;
	LRSETTOOLCORROUT : LREAL;
	XMARKWINDOWTEACHEDTOOL : BOOL;
END_VAR
VAR
	TM_SYNCANDCORRECTIONSTATECONFIG : L_TB2P_ModuleHandlerConfig;
	XTEACHMARKWINDOW_INT : BOOL;
	XTEACHMARKWINDOWTOOL_INT : BOOL;
	XGEARFACTORCORR_INT : BOOL;
	XGEARFACTORCORRHOLD_INT : BOOL;
	XMASTERVALUECORRENABLED_INT : BOOL;
	_LRCORRECTIONDIFF : LREAL;
	_XCORRACTIVE : BOOL;
	LRCORRREGPOSOLD : LREAL;
	FM_L_TS2P_MASTERVALUECORRECTION : L_TS2P_MasterValueCorrection;
	FM_L_TS2P_TOOLCORRECTION : L_TS2P_ToolCorrection;
END_VAR
END_FUNCTION_BLOCK

METHOD CALL_FM_MASTERVALUECORRECTION
END_METHOD

METHOD CALL_FM_MASTERVALUECORRECTION_INPUT
END_METHOD

METHOD CALL_FM_SYNCHRONIZEDDRIVE_INPUT
END_METHOD

METHOD CALL_FM_TOOLCORRECTION : BOOL
END_METHOD

METHOD CALL_FM_TOOLCORRECTION_INPUT : BOOL
END_METHOD

METHOD CALL_ERRORHANDLER
END_METHOD

METHOD CALL_FBMETHODS
END_METHOD

METHOD CALL_INIT_FM
END_METHOD

METHOD CALL_INTERNALCTRL
END_METHOD

METHOD CALL_OUTPUT
END_METHOD

METHOD CALL_OUTPUT_SF
END_METHOD

METHOD CALL_REQUESTS_EXT
END_METHOD

METHOD CALL_RESETCOMMANDS
END_METHOD

METHOD CALL_RESETOUTPUT
END_METHOD

METHOD CALL_STATEMACHINE
END_METHOD

METHOD CALL_S000_CYCLIC
END_METHOD

METHOD CALL_S002_STANDBY
END_METHOD

METHOD CALL_S996_STOP
END_METHOD

METHOD CALL_S999_ERROR
END_METHOD

METHOD CALL_T000_ALLSTATES
END_METHOD

(* ---- L_TS2P_TM_SYNCPOSBASE.fb ---- *)
FUNCTION_BLOCK L_TS2P_TM_SYNCPOSBASE EXTENDS L_TB2M_TM_MotionControl
VAR_INPUT
	MASTERVALUES : L_MC1P_IAXIS_REF_MASTERVALUES;
	XSYNCIN : BOOL;
	XSYNCPOSRESTORE : BOOL;
	LRSETBASEVEL : LREAL;
	LRSETOFFSETPOS : LREAL;
	XTRIMPOS : BOOL;
	XTRIMNEG : BOOL;
	XTRIMRESET : BOOL;
END_VAR
VAR_OUTPUT
	XSYNCHRONISED : BOOL;
	XACCDECSYNC : BOOL;
	XOFFSETTRIMACTIVE : BOOL;
	XBASEVELOCITYACTIVE : BOOL;
	LROFFSETTOTAL : LREAL;
END_VAR
VAR
	TM_SYNCPOS : L_TB2P_ModuleHandlerConfig;
	ITFSYNCPOSBASE : L_TS2P_ISyncPosBase := THIS^;
	SCDATA_INT : L_TS2P_scData_TM_SyncPosBase;
	PDATA : POINTER TO L_TS2P_scData_TM_SyncPosBase := ADR(scData_Int);
	PPAR : POINTER TO L_TS2P_scPar_TM_SyncPosBase;
	PSF : POINTER TO L_TS2P_scSF_TM_SyncPosBase;
	PAP : POINTER TO L_TS2P_scAP_TM_SyncPosBase;
	FB_CONDAXISMOVING : L_TB2P_AxisMoving;
	FB_CONDMASTERDIRECTION : L_TB2P_ConditionMasterDirection;
	FB_CONDBASEVELOCITYDIRECTION : L_TB2P_ConditionBaseVelocityDirection;
	FB_CONDSYNCPARAMETER : L_TS2P_ConditionSyncParameter;
	FB_CONDITIONJOGGINGACTIVE : L_UBUP_ConditionInput;
	FB_CONDCOLLECTSYNCIN : L_UBUP_ConditionCollectionAND := STRUCT(aitfCondition := [fb_ConditionOperationEnabled, fb_ConditionLimiter, fb_CondMasterDirection, fb_CondSyncParameter, fb_ConditionJoggingActive, fb_ConditionAxisNotStopping]);
	FB_CONDCOLLECTBASEVELOCITY : L_UBUP_ConditionCollectionAND := STRUCT(aitfCondition := [fb_CondBaseVelocityDirection, fb_CondCollectOperationEnabledLimiter, fb_ConditionJoggingActive, fb_ConditionAxisNotStopping]);
	FB_TRANSITION2BASEVELOCITYACCDEC : L_UBUP_RequestTransitionLevel;
	FB_TRANSITION2BASEVELOCITY : L_UBUP_RequestTransitionEdge;
	FB_TRANSITION2BASEVELOCITYZERO : L_UBUP_RequestTransitionLevel;
	FB_TRANSITION2SYNCIN : L_UBUP_RequestTransitionLevel;
	FB_TRANSITION2SYNCOUT : L_UBUP_RequestTransitionEdge;
	FB_TRANSITION2SYNCHRONIZED : L_UBUP_RequestTransitionLevel;
	FB_OFFSETANDTRIMX : L_TS2P_OffsetAndTrim;
	FB_ADDOFFSETCYCLICX : L_MC1P_AddOffsetCyclic;
	FB_GEARBOXPOSITION : L_MB1P_GearboxPositionInput;
	FB_AXISCONVERTER : L_MC2P_AxisConverterBase;
	FB_SYNCPOSRESTOREOFFSET : L_TS2P_OffsetAndTrim;
	FB_CLUTCHEXTENDEDBASE : L_TB2P_ClutchExtendedBase;
	FB_ALLOWEDDIRECTION : L_TS2P_AllowedDirection;
	FB_CONTROLSETVALUES : L_MC1P_ControlSetValues;
	MASTERVALUES_INT : L_MC1P_SetAxisRefMasterValues;
	_ITFREQUESTCONDITIONWARNINGHIGHPRIO : L_UBUP_IRequest;
	IVISFRAMESIGNALFLOW : INT;
	DIFRAMESF : DINT;
	CONNECTOR : __SYSTEM.IQueryInterface;
	SYNCPOSBASEEXTENSION : L_TS2P_ISyncPosBase;
END_VAR
END_FUNCTION_BLOCK

METHOD HANDLEREJECTEDREQUEST : BOOL
VAR_INPUT
	ITFREQUESTANNOUNCED : L_UBUP_IRequest;
END_VAR
VAR_OUTPUT
	ITFALTERNATIVEREQUEST : L_UBUP_IRequest;
END_VAR
END_METHOD

METHOD CALLFBS
VAR_INPUT
	ECASE : L_UBUP_StateHandleCase;
END_VAR
END_METHOD

METHOD CALLSTATE
VAR_INPUT
	ITFSTATESERVER : L_UBUP_IStateServer;
	ISTATE : INT;
	ECASE : L_UBUP_StateHandleCase;
END_VAR
END_METHOD

METHOD CHECKTRANSITION
VAR_INPUT
	ITFSTATESERVER : L_UBUP_IStateServer;
END_VAR
END_METHOD

METHOD FINALIZECYCLE
END_METHOD

METHOD PREPARECYCLE
END_METHOD

METHOD SETADDMODULEINFO
VAR_INPUT
	ESUBCOMPTYPE : UDINT;
	SLICINFO : STRING(10);
END_VAR
END_METHOD

METHOD STIMULATETRANSITION
VAR_INPUT
	ECASE : L_UBUP_StateHandleCase;
END_VAR
END_METHOD

METHOD CALL_SETLOCALMASTERVALUES
END_METHOD

METHOD STATE_01_BASEVEL_ACC_DEC
VAR_INPUT
	ECASE : L_UBUP_StateHandleCase;
	ISTATESERVER : L_UBUP_IStateServer;
END_VAR
END_METHOD

METHOD STATE_02_BASEVEL_2_STANDSTILL
VAR_INPUT
	ECASE : L_UBUP_StateHandleCase;
	ISTATESERVER : L_UBUP_IStateServer;
END_VAR
END_METHOD

METHOD STATE_03_BASEVELOCITY
VAR_INPUT
	ECASE : L_UBUP_StateHandleCase;
	ISTATESERVER : L_UBUP_IStateServer;
END_VAR
END_METHOD

METHOD STATE_11_SYNC_ACC
VAR_INPUT
	ECASE : L_UBUP_StateHandleCase;
	ISTATESERVER : L_UBUP_IStateServer;
END_VAR
END_METHOD

METHOD STATE_12_SYNC_DEC
VAR_INPUT
	ECASE : L_UBUP_StateHandleCase;
	ISTATESERVER : L_UBUP_IStateServer;
END_VAR
END_METHOD

METHOD STATE_13_SYNCHRONISED
VAR_INPUT
	ECASE : L_UBUP_StateHandleCase;
	ISTATESERVER : L_UBUP_IStateServer;
END_VAR
END_METHOD

METHOD ADDOFFSET
VAR_INPUT
	ITFTECHMODULE : L_TS2P_ISyncPosBase;
	LRSETPOS : LREAL;
	LRSETVEL : LREAL;
	LRSETOFFSET : LREAL;
	LRSETOFFSETVEL : LREAL;
	ETRAVERSINGRANGE : L_MC1P.L_MC1P_TraversingRange;
	LRCYCLELENGTH : LREAL;
END_VAR
VAR_OUTPUT
	XERROR : BOOL;
	EERRORID : L_IE1P.L_IE1P_Error;
	LRSETPOSOUT : LREAL;
	LRSETVELOUT : LREAL;
END_VAR
END_METHOD

METHOD CLUTCH
VAR_INPUT
	ITFTECHMODULE : L_TS2P_ISyncPosBase;
	XENABLE : BOOL;
	XSYNCIN : BOOL;
	LRSETBASEVELOCITY : LREAL;
	ESYNCMODE : L_TB2P_SyncMode;
	EALLOWEDDIRECTION : L_TB2P_AllowedDirection;
	LRSYNCVEL : LREAL;
	LRSYNCACC : LREAL;
	LRSYNCDEC : LREAL;
	LRSYNCJERK : LREAL;
	LRSYNCINDIST : LREAL;
	LRSYNCOUTDIST : LREAL;
	LRSYNCOUTPOS : LREAL;
	XLOADCLUTCHOFFSET : BOOL;
	LRLOADCLUTCHOFFSET : LREAL;
	LRCYCLICMASTERPOS : LREAL;
	LRCYCLICMASTERVEL : LREAL;
	ETRAVERSINGRANGEMASTER : L_MC1P_TraversingRange;
	LRCYCLELENGTHMASTER : LREAL;
	LRCYCLICAXISPOS : LREAL;
	LRCYCLICAXISVEL : LREAL;
	LRCYCLICAXISACC : LREAL;
	ETRAVERSINGRANGEAXIS : L_MC1P_TraversingRange;
	LRCYCLELENGTHAXIS : LREAL;
END_VAR
VAR_OUTPUT
	XERROR : BOOL;
	EERRORID : L_IE1P.L_IE1P_Error;
	XBUSY : BOOL;
	XDONE : BOOL;
	XSYNCHRONISED : BOOL;
	XACCDECSYNC : BOOL;
	XINBASEVELOCITY : BOOL;
	LRSETPOSOUT : LREAL;
	LRSETVELOUT : LREAL;
	LRSETACCOUT : LREAL;
	LRCLUTCHOFFSETOUT : LREAL;
END_VAR
END_METHOD

METHOD GEARBOX
VAR_INPUT
	ITFTECHMODULE : L_TS2P_ISyncPosBase;
	XENABLE : BOOL;
	LRSETPOSX : LREAL;
	LRSETVELX : LREAL;
	DWNUMERATOR : DWORD;
	DWDENOMINATOR : DWORD;
	LRCYCLELENGTHX : LREAL;
	LRCYCLELENGTHY : LREAL;
	ETRAVERSINGRANGEX : L_MC1P.L_MC1P_TraversingRange;
	ETRAVERSINGRANGEY : L_MC1P.L_MC1P_TraversingRange;
	XLOADGEARBOXPOS : BOOL;
	LRLOADGEARBOXPOS : LREAL;
END_VAR
VAR_OUTPUT
	XERROR : BOOL;
	EERRORID : L_IE1P.L_IE1P_Error;
	LRSETPOSOUT : LREAL;
	LRSETVELOUT : LREAL;
END_VAR
END_METHOD

METHOD OFFSETANDTRIM
VAR_INPUT
	ITFTECHMODULE : L_TS2P_ISyncPosBase;
	XENABLE : BOOL;
	LRSETOFFSET : LREAL;
	XTRIMPOS : BOOL;
	XTRIMNEG : BOOL;
	LRSETTRIMDISTANCE : LREAL;
	ETRIMMODE : L_TS2P_TrimMode;
	XLOADOFFSET : BOOL;
	XRESETTRIMOFFSET : BOOL;
	LRSETVEL : LREAL;
	LRSETACC : LREAL;
	LRSETDEC : LREAL;
	LRSETJERK : LREAL;
	WACTDIRECTION : WORD;
	EALLOWEDDIRECTION : L_TB2P.L_TB2P_AllowedDirection;
	LRCYCMASTERPOS : LREAL;
	LRCYCMASTERVEL : LREAL;
	LRCYCMASTERACC : LREAL;
END_VAR
VAR_OUTPUT
	XERROR : BOOL;
	EERRORID : L_IE1P.L_IE1P_Error;
	XBUSY : BOOL;
	XDONE : BOOL;
	LRSETOFFSETOUTTOTAL : LREAL;
	LRSETOFFSETOUTTOTALVEL : LREAL;
	LRSETOFFSETOUT : LREAL;
	LRSETOFFSETOUTTRIM : LREAL;
END_VAR
END_METHOD

METHOD CALL_ALLOCPOINTADR
END_METHOD

METHOD CALL_EXIT_CALLFBS
END_METHOD

METHOD CALL_INIT_CALLFBS
END_METHOD

METHOD CALL_INTERNALCTRL
END_METHOD

METHOD CALL_RESETOUTPUT
END_METHOD

METHOD MAPTMSTATE
VAR_INPUT
	ETMSTATEINTERNAL : L_TB2P_States;
END_VAR
VAR_OUTPUT
	ETMSTATEEXTERNAL : L_TB2P_States;
END_VAR
END_METHOD

(* ---- L_TS2P_TM_SYNCPOSBASE_V2.fb ---- *)
FUNCTION_BLOCK L_TS2P_TM_SYNCPOSBASE_V2 EXTENDS L_TB2P_SyncMotionControl
VAR_OUTPUT
	PPAR : POINTER TO L_TS2P_scPar_TM_SyncAndCorrectionState := ADR(scPar_int);
	PSF : POINTER TO L_TS2P_scSF_TM_SyncAndCorrectionState;
	PAP : POINTER TO L_TS2P_scAP_TM_SyncAndCorrectionState;
END_VAR
VAR_IN_OUT
	XSYNCIN : BOOL;
	XSYNCPOSRESTORE : BOOL;
	LRSETBASEVEL : LREAL;
	LRSETOFFSETPOS : LREAL;
	XTRIMPOS : BOOL;
	XTRIMNEG : BOOL;
	XTRIMRESET : BOOL;
	SCSIGNALFLOW : L_TS2P_scSF_TM_SyncPosBase;
	XSYNCHRONISED : BOOL;
	XACCDECSYNC : BOOL;
	XOFFSETTRIMACTIVE : BOOL;
	XBASEVELOCITYACTIVE : BOOL;
	LROFFSETTOTAL : LREAL;
END_VAR
VAR
	TM_SYNCPOSBASECONFIG : L_TB2P_ModuleHandlerConfig;
	SCPAR_INT : L_TS2P_scPar_TM_SyncAndCorrectionState;
	XSYNCIN_INT : BOOL;
	XSYNCIN_OLD : BOOL;
	LRSETOFFSETSLAVE_INT : LREAL;
	XTRIMPOS_INT : BOOL;
	XTRIMNEG_INT : BOOL;
	XTRIMRESET_INT : BOOL;
	LRSETOFFSETPOS_INT : REAL;
	LROFFSETTRIM_STORE : LREAL;
	_XSYNCDRIVEENABLE : BOOL;
	_XSYNCDRIVESYNCPOS : BOOL;
	_LRSNYCDRIVESETSLAVEPOSOUT : LREAL;
	_LRSYNCDRIVESETOFFSET : LREAL;
	_LRSYNCDRIVESETOFFSETOUT : LREAL;
	_XLOADSTARTSLAVEPOS : BOOL;
	_LRSTARTSLAVEPOS : LREAL;
	_XLOADGEARBOXPOS : BOOL;
	_LRLOADGEARBOXPOS : LREAL;
	_XLOADOFFSETSYNC : BOOL;
	_LRLOADOFFSETSYNC : LREAL;
	MP03_LRSETGEARBOXPOSOUT : LREAL;
	XLOADTRIMOFFSET : BOOL;
	_LRLOADTRIMOFFSET : LREAL;
	_LRSETTRIMOFFSETOUT : LREAL;
	_LRSETTOTALOFFSETOUT : LREAL;
	_XSYNCDRIVESYNCOUTINSTANT : BOOL;
	_XSYNCDRIVETRIMPOS : BOOL;
	_XSYNCDRIVETRIMNEG : BOOL;
	_XSYNCDRIVESYNCOUTDONE : BOOL;
	_LRSYNCDRIVEOFFSETSYNCPOS : LREAL;
	_XSYNCDRIVESYNCHRONISED : BOOL;
	_XSYNCDRIVETRIMBUSY : BOOL;
	_XSYNCDRIVEACCDECSYNC : BOOL;
	_XSYNCDRIVEACCDECSYNCOLD : BOOL;
	MP04_LRSETCLUTCHPOS : LREAL;
	_XBASEVELSYNCHRONISED : BOOL;
	XINVALIDBASEVELFLAG : BOOL;
	_XLOADOFFSETX : BOOL;
	XSYNCPOSRESTORE_INT : BOOL;
	_XLOADOFFSETMASTER : BOOL;
	LRFACTORMASTERTOSLAVE : LREAL;
	_LRSYNCDRIVESETOFFSETOUTMASTER : LREAL;
	XQSPAPPLICATION_OLD : BOOL;
	LRSETBASEVEL_INT : LREAL;
	_XACCDECSYNC : BOOL;
	XABORTSYNC_INT : BOOL;
	XENABLEAXISCONTROLBYPOS : BOOL;
	IACTMASTERDIRECTIONTMP : INT;
	XWARNINGDIRECTIONDISABLEDSYNCINT : BOOL;
	XWARNINGDIRECTIONDISABLEDBASEVEL : BOOL;
	FM_L_TS2P_SYNCDRIVE : L_TS2P_SyncDrivePos;
	FB_AXISCONTROLBYPOS : L_MC1P_ControlSetValues;
	FB_SETACTUALPOSITION : MC_SetPosition;
	FB_ALLOWEDDIRECTION : L_TS2P_AllowedDirection;
	XSYNCFLAG_INT : BOOL;
	XDESYNCFLAG_INT : BOOL;
	XENABLEOLD : BOOL;
END_VAR
END_FUNCTION_BLOCK

METHOD CALL_FB_ALLOWEDDIRECTION
END_METHOD

METHOD CALL_FM_SYNCHRONIZEDDRIVE
END_METHOD

METHOD CALL_FM_SYNCHRONIZEDDRIVE_INPUT
END_METHOD

METHOD CALL_FM_TOOLCORRECTION : BOOL
END_METHOD

METHOD CALL_FM_TOOLCORRECTION_INPUT : BOOL
END_METHOD

METHOD CALL_ALLOCPOINTADR
END_METHOD

METHOD CALL_AXISCONTROLBYPOS
END_METHOD

METHOD CALL_AXISCONTROLBYPOS_INPUT
END_METHOD

METHOD CALL_CALCFACTORMASTERTOSLAVE
END_METHOD

METHOD CALL_CTRLREQACTIVE : BOOL
END_METHOD

METHOD CALL_ERRORHANDLER
END_METHOD

METHOD CALL_FBMETHODS
END_METHOD

METHOD CALL_INITDONE
END_METHOD

METHOD CALL_INITROUTINE
END_METHOD

METHOD CALL_INIT_FM
END_METHOD

METHOD CALL_INTERNALCTRL
END_METHOD

METHOD CALL_MASTERAXISREF
VAR_INPUT
	MASTERVALUES : L_MC1P_IAXIS_REF_MASTERVALUES;
END_VAR
END_METHOD

METHOD CALL_OUTPUT
END_METHOD

METHOD CALL_OUTPUT_SF
END_METHOD

METHOD CALL_REQUESTS_EXT
END_METHOD

METHOD CALL_RESETCOMMANDS
END_METHOD

METHOD CALL_RESETOUTPUT
END_METHOD

METHOD CALL_STATEMACHINE
END_METHOD

METHOD CALL_ABC_INPUT_PROFILEPARAMETER
END_METHOD

METHOD CALL_S000_CYCLIC
END_METHOD

METHOD CALL_S002_STANDBY
END_METHOD

METHOD CALL_S030_SYNCHRONISING_POS
END_METHOD

METHOD CALL_S031_POS_IS_SYNCHRONISED
END_METHOD

METHOD CALL_S051_BASEVELOCITY
END_METHOD

METHOD CALL_S996_STOP
END_METHOD

METHOD CALL_S999_ERROR
END_METHOD

METHOD CALL_T000_ALLSTATES
END_METHOD

METHOD CALL_T030_DESYNCHRONISING_POS
END_METHOD

METHOD CALL_T030_SYNCHRONISING_POS
END_METHOD

METHOD CALL_T031_POS_IS_SYNCHRONISED
END_METHOD

METHOD CALL_T051_BASEVELOCITY
END_METHOD

METHOD CALL_050_ABORT
END_METHOD

METHOD CALL_S000_CYCLIC_OUT
END_METHOD

METHOD CALL_S003_HOMING_OUT
END_METHOD

METHOD CALL_S010_JOGGING_OUT
END_METHOD

METHOD CALL_S014_MOVEABS_OUT
END_METHOD

METHOD CALL_S015_MOVEREL_OUT
END_METHOD

METHOD CALL_S996_STOP_OUT
END_METHOD

METHOD CALL_S999_ERROR_OUT
END_METHOD

METHOD CALL_STATEMACHINE_OUT
END_METHOD

METHOD CALL_T000_ALLSTATES_OUT
END_METHOD

(* ---- L_TS2P_TOOLCORRECTION.fb ---- *)
FUNCTION_BLOCK L_TS2P_TOOLCORRECTION
VAR_INPUT
	XENABLE : BOOL;
	XACTIVATECORRECTION : BOOL;
	TPRECDATA : L_MC1P_TpReceiveData;
	LRSENSORTOOLDISTANCE : LREAL;
	LRMAXCORRNEG : LREAL;
	LRMAXCORRPOS : LREAL;
	LRUPPERCORRPOS : LREAL;
	LRLOWERCORRPOS : LREAL;
	DNNUMAXISY : DWORD;
	DNDENAXISY : DWORD;
	XENABLEMARKWINDOW : BOOL;
	XTEACHMARKWINDOW : BOOL;
	LRMARKWINDOWSIZE : LREAL;
	LRSETOFFSETMARKWINDOW : LREAL;
	DWMAXNUMBERVIRTUALMARKS : DWORD;
	ECORRMODE : L_TS2P_CorrectionMode;
	LRCORRVEL : LREAL;
	LRCORRACC : LREAL;
	LRCORRDEC : LREAL;
	LRCORRJERK : LREAL;
END_VAR
VAR_OUTPUT
	XERROR : BOOL;
	XWARNING : BOOL;
	EERRORID : WORD;
	XCORRLIMITED : BOOL;
	LRACTMARKERROR : LREAL;
	LRACTMARKDIST : LREAL;
	XINITDONE : BOOL;
	XCORRACTIVE : BOOL;
	XMARKRECEIVED : BOOL;
	LRSENSORACTPOS : LREAL;
	LRSENSORSETPOS : LREAL;
	XMARKWINDOWOPEN : BOOL;
	XMARKOUTOFWINDOW : BOOL;
	XMARKNOTDETECTED : BOOL;
	XMARKWINDOWTEACHED : BOOL;
END_VAR
VAR_IN_OUT
	AXIS : AXIS_REF;
END_VAR
VAR
	SPEEDTOPOSINTEGRATE : L_MC1P_IntegrateAxis;
	TPLIMITDIFF : L_TS2P_TpLimitDiff;
	FB_ADDOFFSET : L_MC1P_AddOffsetCyclic;
	TPCALCDIFF : L_MC1P_TpCalcDiff;
	TP_CONVERTER : L_TB2P_TP_Converter;
	DISTCORRECTIONWINDOW : L_TS2P_DistCorrectionWindow;
	MARKWINDOW : L_TS2P_MarkWindowRelative;
	MARKSTACK : L_TS2P_MarkStack;
	TPVIRTUALACTPOS : L_TS2P_TpVirtualActPos;
	FB_PROFILEGENERATOR : L_MC1P_ProfileGenerator;
	FB_INTEGRATOR : L_MC1P_IntegrateAxis;
	SCPROFILEPARAMETER : L_MC1P_ProfileParameter;
	LRMARKSENSORPOS : LREAL;
	LRGEARINGFAKTOR : LREAL := 1.0;
	XERROR_TM : BOOL;
	EERRORID_TM : L_IE1P_Error;
	LRTPDIFFERENCE : LREAL;
	XLOADMARKSENSORPOS_OLD : BOOL;
	XTPRECEIVED_OLD : BOOL;
	LRMARKWINDOWSIZE_INT : LREAL;
	XTPINWINDOW : BOOL;
	LRPOS_INT : LREAL;
	XTPRECEIVEDOUT_INT : BOOL;
	LRTPACTPOSITION_INT : LREAL;
	LRTPDIFFERENCELIM_INT : LREAL;
	LROFFSETPOSCTRL_INT : LREAL;
	LRPOSOUT_INT : LREAL;
	LRVELOUT_INT : LREAL;
	XCORRACTIVE_INT : BOOL;
	XINIT : BOOL := TRUE;
	XTPCORRECTIONACTIVE : BOOL := FALSE;
	LRTPAXISSETPOS : LREAL;
	LRMARKDIST_INT : LREAL;
	XZERO : BOOL;
	XHOMINGDONE : BOOL;
	XSTARTREFERENCEACTIVE : BOOL;
	XHOMINGACTIVE : BOOL := FALSE;
	XMARKDISTCHANGED : BOOL;
	LRTPACTPOSIN_OLD : LREAL;
	LRTPAXISACTPOS_OLD : LREAL;
	ICOUNTER : INT := 0;
	XFIRSTTOUCHPROBE : BOOL := TRUE;
	LRMARKSTACKLENGTH : LREAL;
	LRTPDIFFERENCELIMITOUT_INT : LREAL;
	XTPRECEIVESTACKOUT_INT : BOOL;
	XTPNOTDETECTED_INT : BOOL;
	XMAXTPNOTDETECTED : BOOL;
	LRGEARFACTORINTEGRATOR : LREAL;
	LRGEARFACTORGAIN : LREAL := 1;
	LRGEARFACTORNUMERATORCORR : LREAL;
	LRGEARFACTORNUMERATORCORRLIMITED : LREAL;
	LRGEARFACTORDENOMINATOR : LREAL;
	LRGEARFACTORNUMERATOR : LREAL;
	LRTOTALSTACKDIFFERENCEOUT_INT : LREAL := 0;
	LCORRECTIONVELIN : LREAL;
	LRSETPOSCORROUT_OLD : LREAL;
	LRDELTAGEARFACTORCORR : LREAL;
	XTPSENSORTEACHEDOLD : BOOL;
	XTPSENSORTEACHEDATLASTMARK : BOOL;
	XCALCMARKDISTINITIALISED : BOOL;
	XTEACHTPSENSOROLD : BOOL;
	LRTPDEADTIMEDIFF : LREAL;
	XTPRECEIVEDOUTOLD_INT : BOOL;
	LRMARKDISTINTEGRATOR : LREAL;
	LRPOSOUTOLD_INT : LREAL;
	LRCORRPOS_INT : LREAL;
	LRCORRPOSOLD_INT : LREAL := 0;
	XENABLEOLD : BOOL;
	TPRECDATAMARKSTACK : L_MC1P_TpReceiveData;
	TPRECDATAMARKWINDOW : L_MC1P_TpReceiveData;
	XTPRECEIVEDINOLD_INT : BOOL;
	XFIRSTVALUESTORED : BOOL;
	LRAXISSETPOSOLD_INT : LREAL;
	LRCORRRESIDUAL : LREAL;
	ECORRECTIONMODEOLD : L_TS2P_CorrectionMode;
	XCORRECTIONBUSY : BOOL;
END_VAR
END_FUNCTION_BLOCK

METHOD CALL_CALCACTMARKDIST
END_METHOD

METHOD CALL_CALCTOOLERROR
END_METHOD

METHOD CALL_CORRECTIONPOS
END_METHOD

METHOD CALL_CORRECTIONPROFILE
END_METHOD

METHOD CALL_ENABLEREGISTERCONTROL
END_METHOD

METHOD CALL_ERRORHANDLER
END_METHOD

METHOD CALL_FB
END_METHOD

METHOD CALL_INPUT
END_METHOD

METHOD CALL_LIMIT
END_METHOD

METHOD CALL_MARKDISTCHANGE
END_METHOD

METHOD CALL_MARKSENSORPOS
END_METHOD

METHOD CALL_MARKSTACK
END_METHOD

METHOD CALL_MARKWINDOW
END_METHOD

METHOD CALL_NOTENABLE
END_METHOD

METHOD CALL_OUTPUT
END_METHOD

METHOD CALL_RESET
END_METHOD

METHOD CALL_RESETOUTPUTS
END_METHOD

METHOD CALL_SETCORRECTION
END_METHOD

METHOD CALL_TPCONVERTER
END_METHOD

METHOD CALL_VIRTUALACTPOS
END_METHOD

METHOD GET_ACTMARKERRORLIMITED : LREAL
END_METHOD

METHOD GET_ACTUALMARKDIST : LREAL
END_METHOD

METHOD GET_CORRREGPOS : LREAL
END_METHOD

METHOD GET_INTEGRATORREGPOS : LREAL
END_METHOD

METHOD GET_MARKERRORUNLIMITED : LREAL
END_METHOD

METHOD GET_MARKPOSITIONINREGISTER : LREAL
END_METHOD

METHOD GET_MARKRECEIVEUNLIMITED : BOOL
END_METHOD

METHOD GET_MARKRECEIVEDLIMITED : BOOL
END_METHOD

METHOD GET_MARKWINDOWCOMP : BOOL
END_METHOD

METHOD GET_REGISTERINPUTVEL : LREAL
END_METHOD

METHOD GET_SETVELOCITYREGISTER : LREAL
END_METHOD

METHOD GET_LRMARKSTACKLENGTH : LREAL
END_METHOD

(* ---- L_TS2P_TPLIMITDIFF.fb ---- *)
FUNCTION_BLOCK L_TS2P_TPLIMITDIFF
VAR_INPUT
	XTPRECEIVED : BOOL;
	LRSETTPDIFFERENCE : LREAL;
	LRSETLIMITMIN : LREAL := -100;
	LRSETLIMITMAX : LREAL := 100;
END_VAR
VAR_OUTPUT
	XTPRECEIVEDOUT : BOOL;
	XLIMITACTIVE : BOOL;
	LRTPDIFFERENCELIM : LREAL;
END_VAR
VAR
	XTPRECEIVEDOLD : BOOL;
	XINITDONE : BOOL;
END_VAR
END_FUNCTION_BLOCK

(* ---- L_TS2P_TPVIRTUALACTPOS.fb ---- *)
FUNCTION_BLOCK L_TS2P_TPVIRTUALACTPOS
VAR_INPUT
	XTPWINDOWOPEN : BOOL;
	XTPRECEIVEDIN : BOOL;
	XMAXTPNOTDETECTED : BOOL;
	LRSETTPPOSIN : LREAL;
	LRACTTPPOSIN : LREAL;
END_VAR
VAR_OUTPUT
	XTPRECEIVEDOUT : BOOL;
	LRACTTPPOS : LREAL;
END_VAR
VAR
	XTPRECEIVEDINOLD : BOOL;
	XFLAGWINDOWOPENANDNOTP : BOOL := FALSE;
	XWINDOWOPENOLD : BOOL;
	XVIRTUALTPACTIVE : BOOL;
END_VAR
END_FUNCTION_BLOCK

(* ---- L_TS2P_VISUPOOL.fb ---- *)
FUNCTION_BLOCK L_TS2P_VISUPOOL
VAR
	M_STNAMESPACE : STRING(80);
	M_STHELPVARID : STRING;
	M_STHELPVARPATH : STRING(255);
	M_STHELP : STRING;
	M_REGISTERIMAGES : BOOL := TRUE;
END_VAR
END_FUNCTION_BLOCK

METHOD FB_INIT : BOOL
VAR_INPUT
	BINITRETAINS : BOOL;
	BINCOPYCODE : BOOL;
END_VAR
END_METHOD

METHOD FB_REINIT : BOOL
END_METHOD

METHOD FB_EXIT : BOOL
VAR_INPUT
	BINCOPYCODE : BOOL;
END_VAR
END_METHOD

(* ---- L_TT1P_INPOSITION.fb ---- *)
FUNCTION_BLOCK L_TT1P_INPOSITION
VAR_INPUT
	XENABLE : BOOL;
	LRPOSWINDOW : LREAL;
	LRPOSTIME : LREAL;
	XHOLDSETPOS : BOOL;
END_VAR
VAR_OUTPUT
	XINPOSITION : BOOL;
	XBUSY : BOOL;
	LRHOLDPOSITION : LREAL;
	XERROR : BOOL;
	EERRORID : L_IE1P_Error;
END_VAR
VAR_IN_OUT
	AXIS : AXIS_REF;
END_VAR
VAR
	XINTOL : BOOL;
	XENABLEOLD : BOOL := FALSE;
	XHOLDSETPOSOLD : BOOL := FALSE;
	LRSETPOSITIONOLD : LREAL;
	XSETPOSITIONCHG : BOOL;
	INPOSITION_TON : TON;
	INPOSITION_F_TRIG : F_TRIG;
	TIMEOUT_TON : TON;
END_VAR
END_FUNCTION_BLOCK

METHOD FB_RESET : BOOL
END_METHOD
